(* CODESYS project beveling.project

Project tree, tasks and I/O mapping:
  Device : AM523-0808TN, Shenzhen Inovance Control Technology, version 3.5.11.50
      settings: PersistentStartAdddr = 0; PersistentStartEndAddr = 524287; Mode = 1
    application Application
      libraries: Standard, * (System); CmpEventMgr, 3.5.8.0 (System); Component Manager, 3.5.9.0 (System); CmpApp, 3.5.11.0 (System); CmpIecTask, 3.5.9.0 (System); CmpHCMotion, 1.1.8.0 (Inovance)
      task MainTask (cyclic, interval 4 ms, priority 1) calls nothing
      task ETHERCAT1 (cyclic, interval 2000 µs, priority 0) calls ETHERCAT1.EtherCAT_Task, PLC_PRG
      01_Data/
        global variables GVL_Parameters
        global variables GVL_IO_Physical
        global variables GVL_Modbus
        global variables GVL_RealDevice
        global variables GVL_DeviceIds
        global variables GVL_Simulation
        global variables GVL_Interface
        global variables GVL_IO
      06_Simulation/
        function block FB_SimDevice [ST]
        function block FB_SimPlant [ST]
      program PLC_PRG [ST]
      global variables GVL_Motion
      04_Machine/
        function block FB_IOMap [ST]
        function block FB_AlarmManager [ST]
        function block FB_PanelInput [ST]
        function block FB_AutoCycle [ST]
        function block FB_Interlocks [ST]
        function F_RecipeValid [ST]
        function block FB_ManualControl [ST]
        function block FB_Machine [ST]
        function block FB_Indicator [ST]
      00_Types/
        data type ST_RealDeviceSettings
        data type ST_MachineStatus
        data type E_MachineMode
        data type ST_Recipe
        data type ST_DeviceStatus
        data type E_DeviceAction
        data type E_MachineState
        data type ST_DeviceCommand
        data type ST_OperatorCommand
        data type ST_DeviceConfig
        data type ST_SimulationSettings
        data type E_DeviceKind
        data type ST_ManualCommand
        data type E_AutoStep
        data type ST_RemoteCommand
        data type ST_PanelInputs
      90_Legacy/
        program PRG_AxisDemo [ST]
      TaskEventPreStart
      05_Communication/
        function block FB_ModbusInterface [ST]
      03_Units/
        function block FB_ReturnKnife [ST]
        function block FB_PostCut [ST]
        function block FB_ResetLength [ST]
        function block FB_Initialize [ST]
        function block FB_Unload [ST]
        function block FB_ClearLength [ST]
        function block FB_ClearanceUnit [ST]
        function block FB_ClearTransfer [ST]
      DifferentialMonitor
      02_Devices/
        function block FB_RealAxis [ST]
        function block FB_RealCylinder [ST]
        function block FB_Motor [ST]
        function block FB_RealCylinderGroup [ST]
        function F_Done [ST]
        function block FB_Valve [ST]
        function F_At [ST]
        function block FB_Axis [ST]
        function F_SafetyBypassActive [ST]
        function block FB_RealSensor [ST]
        function block FB_Cylinder [ST]
        function F_Command [ST]
        function F_NextID [ST]
        function block FB_DeviceManager [ST]
    Device Diagnosis
    HardWare Configuration
    ConfigStorage
    Network Configuration
      LocalBus Config
      EtherCAT Config
    Resources List
    Serial : 串行接口, 汇川技术股份有限公司, version 00.00.00.10
      COM : Serial Port, Inovance, version 00.00.00.10
          settings: Device = AM523-0808TN; devGuid = 'e48f0cf2-85a4-455f-a8e7-135d3403221f'
    Local Bus
      GL20_0032ETN : GL20(GL20S) 32点DO模块, Inovance, version 00.00.00.10
          settings: ModuleBaseInfoStruct.BusType = 10; ModuleBaseInfoStruct.RackNumber = 1; ModuleBaseInfoStruct.SlotNumber = 2
          output Application.xDoG9Valve : BOOL  // QB(I).Q0
          output Application.xDoG1ValveL : BOOL  // QB(I).Q1
          output Application.xDoG1ValveR : BOOL  // QB(I).Q2
          output Application.xDoLampGreen : BOOL  // QB(II).Q0
          output Application.xDoLampRed : BOOL  // QB(II).Q1
          unmapped channels: QB(I), QB(II), QB(III), QB(IV)
      GL20_3200END : GL20(GL20S) 32通道DI模块, Inovance, version 00.00.00.10
          settings: ModuleBaseInfoStruct.BusType = 10; ModuleBaseInfoStruct.RackNumber = 1; ModuleBaseInfoStruct.SlotNumber = 1
          input  Application.xDiG1LRetract : BOOL  // IB(I).I0
          input  Application.xDiG1LExtend : BOOL  // IB(I).I1
          input  Application.xDiG1RRetract : BOOL  // IB(I).I2
          input  Application.xDiG1RExtend : BOOL  // IB(I).I3
          input  Application.xDiG9Retract : BOOL  // IB(I).I4
          input  Application.xDiG9Extend : BOOL  // IB(I).I5
          input  Application.xDiEStop : BOOL  // IB(II).I0
          input  Application.xDiPanelRunStop : BOOL  // IB(II).I1
          input  Application.xDiPanelStart : BOOL  // IB(II).I2
          input  Application.xDiPanelReset : BOOL  // IB(II).I3
          input  Application.xDiPanelInit : BOOL  // IB(II).I4
          input  Application.xDiPanelRunStart : BOOL  // IB(II).I5
          input  Application.xDiPanelAutoMode : BOOL  // IB(II).I6
          input  Application.xDiPanelSafetyPermit : BOOL  // IB(II).I7
          input  Application.xDiMaterialLength : BOOL  // IB(III).I0
          unmapped channels: IB(I), IB(II), IB(III), IB(IV)
    EXP_A : 扩展卡, 汇川技术股份有限公司, version 00.00.00.10
    ETHERCAT1 : EtherCAT Master SoftMotion, 3S - Smart Software Solutions GmbH, version 3.5.11.10
        settings:  = 0; MasterCycleTime = 2000; NetworkName = 'eth1'; SelectNetworkByName = TRUE; DisableTaskGeneration = True; SlaveArrayName = ADR(_EC1_Node)
      ASDA_B3_E_CoE_Drive_4 : Delta ASDA-B3-E EtherCAT(CoE) Drive, Delta Electronics, Inc., order no. ASDA-B3-E CoE Drive, version Revision=16#00030000
          settings: StationAlias = 0; Ring of slave = 0; Configuration address of the slave = 5; DC sync0 cycletime = 2000; DC sync1 cycletime = 2000; Interpolation time period.Value = 2
          unmapped channels: Control Word, Target Position, Target Velocity, Target Torque, Touch Probe Function, Status Word, Actual Position, Velocity actual value, Actual Torque, Touch Probe Status, Touch Probe Pos1 Pos Value, Digital inputs
        cetui : Axis, Inovance, order no. 0, version 4.0.0.0
            settings: wDriveID = 5; dwRatioTechUnitsDenom = 8388608; iRatioTechUnitsNum = 5; HomingMode = 2; ZeroSignal = 0; StartDirction = -1; EndDirection = -1; PosLimitMode = 1; NegLimitMode = 1; HomingVelocity = 30; HomingApproachVelocity = 10; HomingAcceleration = 100; HomingDeceleration = 100; HomingJerk = 0; HomeMaskDistance = 0; HomePositionOffset = 0; HomePushTime = 0; HomeCompensation = 0; HomeTimeout = 0; HomeCompensationVelocity = 1000; 4000 = 1; 4001 = 1; ScalingIncs = 16777216; ScalingGearOutput1 = 10; 6005 = 1; AdrOffset_8010 = 72; BitOffset_8010 = 0; BitLength_8010 = 16; Address_8010 = '%QW36'; Type_8010 = 'UINT'; AddressPointer_8010 = ADR(%QW36); AdrOffset_8020 = 76; BitOffset_8020 = 0; BitLength_8020 = 32; Address_8020 = '%QD19'; Type_8020 = 'DINT'; AddressPointer_8020 = ADR(%QD19); AdrOffset_8030 = 80; BitOffset_8030 = 0; BitLength_8030 = 32;
              Address_8030 = '%QD20'; Type_8030 = 'DINT'; AddressPointer_8030 = ADR(%QD20); AdrOffset_8040 = 84; BitOffset_8040 = 0; BitLength_8040 = 16; Address_8040 = '%QW42'; Type_8040 = 'INT'; AddressPointer_8040 = ADR(%QW42); AdrOffset_8050 = 4294967295; BitOffset_8050 = 0; BitLength_8050 = 0; Address_8050 = ''; Type_8050 = ''; AddressPointer_8050 = 0; AdrOffset_8060 = 86; BitOffset_8060 = 0; BitLength_8060 = 16; Address_8060 = '%QW43'; Type_8060 = 'UINT'; AddressPointer_8060 = ADR(%QW43); AdrOffset_8070 = 4294967295; BitOffset_8070 = 0; BitLength_8070 = 0; Address_8070 = ''; Type_8070 = ''; AddressPointer_8070 = 0; AdrOffset_8080 = 4294967295; BitOffset_8080 = 0; BitLength_8080 = 0; Address_8080 = ''; Type_8080 = ''; AddressPointer_8080 = 0; AdrOffset_8090 = 4294967295; BitOffset_8090 = 0; BitLength_8090 = 0; Address_8090 = ''; Type_8090 = ''; AddressPointer_8090 = 0; AdrOffset_8100 = 4294967295;
              BitOffset_8100 = 0; BitLength_8100 = 0; Address_8100 = ''; Type_8100 = ''; AddressPointer_8100 = 0; AdrOffset_8510 = 104; BitOffset_8510 = 0; BitLength_8510 = 16; Address_8510 = '%IW52'; Type_8510 = 'UINT'; AddressPointer_8510 = ADR(%IW52); AdrOffset_8520 = 108; BitOffset_8520 = 0; BitLength_8520 = 32; Address_8520 = '%ID27'; Type_8520 = 'DINT'; AddressPointer_8520 = ADR(%ID27); AdrOffset_8530 = 112; BitOffset_8530 = 0; BitLength_8530 = 32; Address_8530 = '%ID28'; Type_8530 = 'DINT'; AddressPointer_8530 = ADR(%ID28); AdrOffset_8540 = 116; BitOffset_8540 = 0; BitLength_8540 = 16; Address_8540 = '%IW58'; Type_8540 = 'INT'; AddressPointer_8540 = ADR(%IW58); AdrOffset_8550 = 4294967295; BitOffset_8550 = 0; BitLength_8550 = 0; Address_8550 = ''; Type_8550 = ''; AddressPointer_8550 = 0; AdrOffset_8560 = 124; BitOffset_8560 = 0; BitLength_8560 = 32; Address_8560 = '%ID31'; Type_8560 = 'UDINT';
              AddressPointer_8560 = ADR(%ID31); AdrOffset_8570 = 118; BitOffset_8570 = 0; BitLength_8570 = 16; Address_8570 = '%IW59'; Type_8570 = 'UINT'; AddressPointer_8570 = ADR(%IW59); AdrOffset_8580 = 120; BitOffset_8580 = 0; BitLength_8580 = 32; Address_8580 = '%ID30'; Type_8580 = 'DINT'; AddressPointer_8580 = ADR(%ID30); AdrOffset_8590 = 4294967295; BitOffset_8590 = 0; BitLength_8590 = 0; Address_8590 = ''; Type_8590 = ''; AddressPointer_8590 = 0; AdrOffset_8600 = 4294967295; BitOffset_8600 = 0; BitLength_8600 = 0; Address_8600 = ''; Type_8600 = ''; AddressPointer_8600 = 0; AdrOffset_8600 = 4294967295; BitOffset_8600 = 0; BitLength_8600 = 0; Address_8610 = ''; Type_8610 = ''; AddressPointer_8610 = 0; AdrOffset_8620 = 4294967295; BitOffset_8620 = 0; BitLength_8620 = 0; Address_8620 = ''; Type_8620 = ''; AddressPointer_8620 = 0; IsValid = True; AxisNumber = 5; IsHostHoming = True;
              PulseSelectIndex = 0
      DM3B_EC542 : DM3B-EC542(COE), Leadshine Technology Co.,Ltd., order no. DM3B-EC542, version Revision=16#00000001
          settings: StationAlias = 0; Ring of slave = 0; Configuration address of the slave = 8; DC sync0 cycletime = 2000; DC sync1 cycletime = 2000
          unmapped channels: Control Word, Profile Target Position, Touch Probe Function, Last Error Code, Status Word, Modes of Operation display, Position Actual Value, Touch Probe Status, Touch Probe 1 Positive Value, Digital Inputs
        dingchang_shangxia : Axis, Inovance, order no. 0, version 4.0.0.0
            settings: wDriveID = 8; dwRatioTechUnitsDenom = 10000; HomingMode = 7; ZeroSignal = 0; StartDirction = -1; EndDirection = 1; PosLimitMode = 0; NegLimitMode = 0; HomingVelocity = 5; HomingApproachVelocity = 2; HomingAcceleration = 100; HomingDeceleration = 100; HomingJerk = 0; HomeMaskDistance = 0; HomePositionOffset = 0; HomePushTime = 0; HomeCompensation = 0; HomeTimeout = 0; HomeCompensationVelocity = 1000; 4000 = 1; 4001 = 0; ScalingIncs = 10000; 6005 = 1; AdrOffset_8010 = 116; BitOffset_8010 = 0; BitLength_8010 = 16; Address_8010 = '%QW58'; Type_8010 = 'UINT'; AddressPointer_8010 = ADR(%QW58); AdrOffset_8020 = 120; BitOffset_8020 = 0; BitLength_8020 = 32; Address_8020 = '%QD30'; Type_8020 = 'DINT'; AddressPointer_8020 = ADR(%QD30); AdrOffset_8030 = 4294967295; BitOffset_8030 = 0; BitLength_8030 = 0; Address_8030 = ''; Type_8030 = '';
              AddressPointer_8030 = 0; AdrOffset_8040 = 4294967295; BitOffset_8040 = 0; BitLength_8040 = 0; Address_8040 = ''; Type_8040 = ''; AddressPointer_8040 = 0; AdrOffset_8050 = 4294967295; BitOffset_8050 = 0; BitLength_8050 = 0; Address_8050 = ''; Type_8050 = ''; AddressPointer_8050 = 0; AdrOffset_8060 = 124; BitOffset_8060 = 0; BitLength_8060 = 16; Address_8060 = '%QW62'; Type_8060 = 'UINT'; AddressPointer_8060 = ADR(%QW62); AdrOffset_8070 = 4294967295; BitOffset_8070 = 0; BitLength_8070 = 0; Address_8070 = ''; Type_8070 = ''; AddressPointer_8070 = 0; AdrOffset_8080 = 4294967295; BitOffset_8080 = 0; BitLength_8080 = 0; Address_8080 = ''; Type_8080 = ''; AddressPointer_8080 = 0; AdrOffset_8090 = 4294967295; BitOffset_8090 = 0; BitLength_8090 = 0; Address_8090 = ''; Type_8090 = ''; AddressPointer_8090 = 0; AdrOffset_8100 = 4294967295; BitOffset_8100 = 0; BitLength_8100 = 0;
              Address_8100 = ''; Type_8100 = ''; AddressPointer_8100 = 0; AdrOffset_8510 = 186; BitOffset_8510 = 0; BitLength_8510 = 16; Address_8510 = '%IW93'; Type_8510 = 'UINT'; AddressPointer_8510 = ADR(%IW93); AdrOffset_8520 = 192; BitOffset_8520 = 0; BitLength_8520 = 32; Address_8520 = '%ID48'; Type_8520 = 'DINT'; AddressPointer_8520 = ADR(%ID48); AdrOffset_8530 = 4294967295; BitOffset_8530 = 0; BitLength_8530 = 0; Address_8530 = ''; Type_8530 = ''; AddressPointer_8530 = 0; AdrOffset_8540 = 4294967295; BitOffset_8540 = 0; BitLength_8540 = 0; Address_8540 = ''; Type_8540 = ''; AddressPointer_8540 = 0; AdrOffset_8550 = 188; BitOffset_8550 = 0; BitLength_8550 = 8; Address_8550 = '%IB188'; Type_8550 = 'SINT'; AddressPointer_8550 = ADR(%IB188); AdrOffset_8560 = 204; BitOffset_8560 = 0; BitLength_8560 = 32; Address_8560 = '%ID51'; Type_8560 = 'UDINT'; AddressPointer_8560 = ADR(%ID51); AdrOffset_8570 = 196;
              BitOffset_8570 = 0; BitLength_8570 = 16; Address_8570 = '%IW98'; Type_8570 = 'UINT'; AddressPointer_8570 = ADR(%IW98); AdrOffset_8580 = 200; BitOffset_8580 = 0; BitLength_8580 = 32; Address_8580 = '%ID50'; Type_8580 = 'DINT'; AddressPointer_8580 = ADR(%ID50); AdrOffset_8590 = 4294967295; BitOffset_8590 = 0; BitLength_8590 = 0; Address_8590 = ''; Type_8590 = ''; AddressPointer_8590 = 0; AdrOffset_8600 = 4294967295; BitOffset_8600 = 0; BitLength_8600 = 0; Address_8600 = ''; Type_8600 = ''; AddressPointer_8600 = 0; AdrOffset_8600 = 4294967295; BitOffset_8600 = 0; BitLength_8600 = 0; Address_8610 = ''; Type_8610 = ''; AddressPointer_8610 = 0; AdrOffset_8620 = 184; BitOffset_8620 = 0; BitLength_8620 = 16; Address_8620 = '%IW92'; Type_8620 = 'UINT'; AddressPointer_8620 = ADR(%IW92); IsValid = True; AxisNumber = 8; IsHostHoming = True; PulseSelectIndex = 0
      ASDA_B3_E_CoE_Drive_1 : Delta ASDA-B3-E EtherCAT(CoE) Drive, Delta Electronics, Inc., order no. ASDA-B3-E CoE Drive, version Revision=16#00030000
          settings: StationAlias = 0; Ring of slave = 0; Configuration address of the slave = 1; DC sync0 cycletime = 2000; DC sync1 cycletime = 2000; Interpolation time period.Value = 2
          unmapped channels: Control Word, Target Position, Target Velocity, Target Torque, Touch Probe Function, Status Word, Actual Position, Velocity actual value, Actual Torque, Touch Probe Status, Touch Probe Pos1 Pos Value, Digital inputs
        qiege : Axis, Inovance, order no. 0, version 4.0.0.0
            settings: wDriveID = 2; dwRatioTechUnitsDenom = 4194304; iRatioTechUnitsNum = 5; HomingMode = 2; ZeroSignal = 0; StartDirction = -1; EndDirection = -1; PosLimitMode = 1; NegLimitMode = 1; HomingVelocity = 40; HomingApproachVelocity = 2; HomingAcceleration = 100; HomingDeceleration = 200; HomingJerk = 0; HomeMaskDistance = 0; HomePositionOffset = 0; HomePushTime = 0; HomeCompensation = 0; HomeTimeout = 0; HomeCompensationVelocity = 1000; 4000 = 1; 4001 = 1; ScalingIncs = 16777216; ScalingMotorTurns2 = 12; 6005 = 240; AdrOffset_8010 = 8; BitOffset_8010 = 0; BitLength_8010 = 16; Address_8010 = '%QW4'; Type_8010 = 'UINT'; AddressPointer_8010 = ADR(%QW4); AdrOffset_8020 = 12; BitOffset_8020 = 0; BitLength_8020 = 32; Address_8020 = '%QD3'; Type_8020 = 'DINT'; AddressPointer_8020 = ADR(%QD3); AdrOffset_8030 = 16; BitOffset_8030 = 0; BitLength_8030 = 32;
              Address_8030 = '%QD4'; Type_8030 = 'DINT'; AddressPointer_8030 = ADR(%QD4); AdrOffset_8040 = 20; BitOffset_8040 = 0; BitLength_8040 = 16; Address_8040 = '%QW10'; Type_8040 = 'INT'; AddressPointer_8040 = ADR(%QW10); AdrOffset_8050 = 4294967295; BitOffset_8050 = 0; BitLength_8050 = 0; Address_8050 = ''; Type_8050 = ''; AddressPointer_8050 = 0; AdrOffset_8060 = 22; BitOffset_8060 = 0; BitLength_8060 = 16; Address_8060 = '%QW11'; Type_8060 = 'UINT'; AddressPointer_8060 = ADR(%QW11); AdrOffset_8070 = 4294967295; BitOffset_8070 = 0; BitLength_8070 = 0; Address_8070 = ''; Type_8070 = ''; AddressPointer_8070 = 0; AdrOffset_8080 = 4294967295; BitOffset_8080 = 0; BitLength_8080 = 0; Address_8080 = ''; Type_8080 = ''; AddressPointer_8080 = 0; AdrOffset_8090 = 4294967295; BitOffset_8090 = 0; BitLength_8090 = 0; Address_8090 = ''; Type_8090 = ''; AddressPointer_8090 = 0; AdrOffset_8100 = 4294967295;
              BitOffset_8100 = 0; BitLength_8100 = 0; Address_8100 = ''; Type_8100 = ''; AddressPointer_8100 = 0; AdrOffset_8510 = 8; BitOffset_8510 = 0; BitLength_8510 = 16; Address_8510 = '%IW4'; Type_8510 = 'UINT'; AddressPointer_8510 = ADR(%IW4); AdrOffset_8520 = 12; BitOffset_8520 = 0; BitLength_8520 = 32; Address_8520 = '%ID3'; Type_8520 = 'DINT'; AddressPointer_8520 = ADR(%ID3); AdrOffset_8530 = 16; BitOffset_8530 = 0; BitLength_8530 = 32; Address_8530 = '%ID4'; Type_8530 = 'DINT'; AddressPointer_8530 = ADR(%ID4); AdrOffset_8540 = 20; BitOffset_8540 = 0; BitLength_8540 = 16; Address_8540 = '%IW10'; Type_8540 = 'INT'; AddressPointer_8540 = ADR(%IW10); AdrOffset_8550 = 4294967295; BitOffset_8550 = 0; BitLength_8550 = 0; Address_8550 = ''; Type_8550 = ''; AddressPointer_8550 = 0; AdrOffset_8560 = 28; BitOffset_8560 = 0; BitLength_8560 = 32; Address_8560 = '%ID7'; Type_8560 = 'UDINT';
              AddressPointer_8560 = ADR(%ID7); AdrOffset_8570 = 22; BitOffset_8570 = 0; BitLength_8570 = 16; Address_8570 = '%IW11'; Type_8570 = 'UINT'; AddressPointer_8570 = ADR(%IW11); AdrOffset_8580 = 24; BitOffset_8580 = 0; BitLength_8580 = 32; Address_8580 = '%ID6'; Type_8580 = 'DINT'; AddressPointer_8580 = ADR(%ID6); AdrOffset_8590 = 4294967295; BitOffset_8590 = 0; BitLength_8590 = 0; Address_8590 = ''; Type_8590 = ''; AddressPointer_8590 = 0; AdrOffset_8600 = 4294967295; BitOffset_8600 = 0; BitLength_8600 = 0; Address_8600 = ''; Type_8600 = ''; AddressPointer_8600 = 0; AdrOffset_8600 = 4294967295; BitOffset_8600 = 0; BitLength_8600 = 0; Address_8610 = ''; Type_8610 = ''; AddressPointer_8610 = 0; AdrOffset_8620 = 4294967295; BitOffset_8620 = 0; BitLength_8620 = 0; Address_8620 = ''; Type_8620 = ''; AddressPointer_8620 = 0; IsValid = True; AxisNumber = 1; IsHostHoming = True;
              PulseSelectIndex = 0
      ASDA_B3_E_CoE_Drive_5 : Delta ASDA-B3-E EtherCAT(CoE) Drive, Delta Electronics, Inc., order no. ASDA-B3-E CoE Drive, version Revision=16#00030000
          settings: StationAlias = 0; Ring of slave = 0; Configuration address of the slave = 7; DC sync0 cycletime = 2000; DC sync1 cycletime = 2000; Interpolation time period.Value = 2
          unmapped channels: Control Word, Target Position, Target Velocity, Target Torque, Touch Probe Function, Status Word, Actual Position, Velocity actual value, Actual Torque, Touch Probe Status, Touch Probe Pos1 Pos Value, Digital inputs
        jixieshou : Axis, Inovance, order no. 0, version 4.0.0.0
            settings: wDriveID = 7; dwRatioTechUnitsDenom = 10485760; HomingMode = 10; ZeroSignal = 0; StartDirction = 1; EndDirection = 1; PosLimitMode = 0; NegLimitMode = 0; HomingVelocity = 10; HomingApproachVelocity = 2; HomingAcceleration = 100; HomingDeceleration = 100; HomingJerk = 0; HomeMaskDistance = 0; HomePositionOffset = 0; HomePushTime = 0; HomeCompensation = 0; HomeTimeout = 0; HomeCompensationVelocity = 1000; 4000 = 1; 4001 = 1; ScalingIncs = 16777216; ScalingMotorTurns2 = 10; ScalingGearOutput1 = 16; 6005 = 1; AdrOffset_8010 = 100; BitOffset_8010 = 0; BitLength_8010 = 16; Address_8010 = '%QW50'; Type_8010 = 'UINT'; AddressPointer_8010 = ADR(%QW50); AdrOffset_8020 = 104; BitOffset_8020 = 0; BitLength_8020 = 32; Address_8020 = '%QD26'; Type_8020 = 'DINT'; AddressPointer_8020 = ADR(%QD26); AdrOffset_8030 = 108; BitOffset_8030 = 0; BitLength_8030 = 32;
              Address_8030 = '%QD27'; Type_8030 = 'DINT'; AddressPointer_8030 = ADR(%QD27); AdrOffset_8040 = 112; BitOffset_8040 = 0; BitLength_8040 = 16; Address_8040 = '%QW56'; Type_8040 = 'INT'; AddressPointer_8040 = ADR(%QW56); AdrOffset_8050 = 4294967295; BitOffset_8050 = 0; BitLength_8050 = 0; Address_8050 = ''; Type_8050 = ''; AddressPointer_8050 = 0; AdrOffset_8060 = 114; BitOffset_8060 = 0; BitLength_8060 = 16; Address_8060 = '%QW57'; Type_8060 = 'UINT'; AddressPointer_8060 = ADR(%QW57); AdrOffset_8070 = 4294967295; BitOffset_8070 = 0; BitLength_8070 = 0; Address_8070 = ''; Type_8070 = ''; AddressPointer_8070 = 0; AdrOffset_8080 = 4294967295; BitOffset_8080 = 0; BitLength_8080 = 0; Address_8080 = ''; Type_8080 = ''; AddressPointer_8080 = 0; AdrOffset_8090 = 4294967295; BitOffset_8090 = 0; BitLength_8090 = 0; Address_8090 = ''; Type_8090 = ''; AddressPointer_8090 = 0; AdrOffset_8100 = 4294967295;
              BitOffset_8100 = 0; BitLength_8100 = 0; Address_8100 = ''; Type_8100 = ''; AddressPointer_8100 = 0; AdrOffset_8510 = 160; BitOffset_8510 = 0; BitLength_8510 = 16; Address_8510 = '%IW80'; Type_8510 = 'UINT'; AddressPointer_8510 = ADR(%IW80); AdrOffset_8520 = 164; BitOffset_8520 = 0; BitLength_8520 = 32; Address_8520 = '%ID41'; Type_8520 = 'DINT'; AddressPointer_8520 = ADR(%ID41); AdrOffset_8530 = 168; BitOffset_8530 = 0; BitLength_8530 = 32; Address_8530 = '%ID42'; Type_8530 = 'DINT'; AddressPointer_8530 = ADR(%ID42); AdrOffset_8540 = 172; BitOffset_8540 = 0; BitLength_8540 = 16; Address_8540 = '%IW86'; Type_8540 = 'INT'; AddressPointer_8540 = ADR(%IW86); AdrOffset_8550 = 4294967295; BitOffset_8550 = 0; BitLength_8550 = 0; Address_8550 = ''; Type_8550 = ''; AddressPointer_8550 = 0; AdrOffset_8560 = 180; BitOffset_8560 = 0; BitLength_8560 = 32; Address_8560 = '%ID45'; Type_8560 = 'UDINT';
              AddressPointer_8560 = ADR(%ID45); AdrOffset_8570 = 174; BitOffset_8570 = 0; BitLength_8570 = 16; Address_8570 = '%IW87'; Type_8570 = 'UINT'; AddressPointer_8570 = ADR(%IW87); AdrOffset_8580 = 176; BitOffset_8580 = 0; BitLength_8580 = 32; Address_8580 = '%ID44'; Type_8580 = 'DINT'; AddressPointer_8580 = ADR(%ID44); AdrOffset_8590 = 4294967295; BitOffset_8590 = 0; BitLength_8590 = 0; Address_8590 = ''; Type_8590 = ''; AddressPointer_8590 = 0; AdrOffset_8600 = 4294967295; BitOffset_8600 = 0; BitLength_8600 = 0; Address_8600 = ''; Type_8600 = ''; AddressPointer_8600 = 0; AdrOffset_8600 = 4294967295; BitOffset_8600 = 0; BitLength_8600 = 0; Address_8610 = ''; Type_8610 = ''; AddressPointer_8610 = 0; AdrOffset_8620 = 4294967295; BitOffset_8620 = 0; BitLength_8620 = 0; Address_8620 = ''; Type_8620 = ''; AddressPointer_8620 = 0; IsValid = True; AxisNumber = 7; IsHostHoming = True;
              PulseSelectIndex = 0
      ASDA_B3_E_CoE_Drive : Delta ASDA-B3-E EtherCAT(CoE) Drive, Delta Electronics, Inc., order no. ASDA-B3-E CoE Drive, version Revision=16#00030000
          settings: StationAlias = 0; Ring of slave = 0; Configuration address of the slave = 2; AutoUpdate = False; DC sync0 cycletime = 2000; DC sync0 cycletime = 2000000; DC sync1 cycletime = 2000; DC sync1 cycletime = 2000000; DC sync1 factor = 'x 1'; Interpolation time period.Value = 2
          unmapped channels: Control Word, Target Position, Target Velocity, Target Torque, Touch Probe Function, Status Word, Actual Position, Velocity actual value, Actual Torque, Touch Probe Status, Touch Probe Pos1 Pos Value, Digital inputs
        xuanzhuan : Axis, Inovance, order no. 0, version 4.0.0.0
            settings: dwRatioTechUnitsDenom = 45088768; iRatioTechUnitsNum = 9; iMovementType = 0; fSWMaxVelocity = 10; fSWMaxAcceleration = 100; fSWMaxDeceleration = 100; HomingMode = 2; ZeroSignal = 0; StartDirction = -1; EndDirection = -1; PosLimitMode = 1; NegLimitMode = 1; HomingVelocity = 3; HomingApproachVelocity = 1; HomingAcceleration = 100; HomingDeceleration = 100; HomingJerk = 0; HomeMaskDistance = 0; HomePositionOffset = 0; HomePushTime = 0; HomeCompensation = 0; HomeTimeout = 0; HomeCompensationVelocity = 1000; 4000 = 4; 4001 = 1; ScalingIncs = 16777216; ScalingMotorTurns2 = 215; ScalingGearOutput1 = 2; 6005 = 360; AdrOffset_8010 = 24; BitOffset_8010 = 0; BitLength_8010 = 16; Address_8010 = '%QW12'; Type_8010 = 'UINT'; AddressPointer_8010 = ADR(%QW12); AdrOffset_8020 = 28; BitOffset_8020 = 0; BitLength_8020 = 32; Address_8020 = '%QD7'; Type_8020 = 'DINT';
              AddressPointer_8020 = ADR(%QD7); AdrOffset_8030 = 32; BitOffset_8030 = 0; BitLength_8030 = 32; Address_8030 = '%QD8'; Type_8030 = 'DINT'; AddressPointer_8030 = ADR(%QD8); AdrOffset_8040 = 36; BitOffset_8040 = 0; BitLength_8040 = 16; Address_8040 = '%QW18'; Type_8040 = 'INT'; AddressPointer_8040 = ADR(%QW18); AdrOffset_8050 = 4294967295; BitOffset_8050 = 0; BitLength_8050 = 0; Address_8050 = ''; Type_8050 = ''; AddressPointer_8050 = 0; AdrOffset_8060 = 38; BitOffset_8060 = 0; BitLength_8060 = 16; Address_8060 = '%QW19'; Type_8060 = 'UINT'; AddressPointer_8060 = ADR(%QW19); AdrOffset_8070 = 4294967295; BitOffset_8070 = 0; BitLength_8070 = 0; Address_8070 = ''; Type_8070 = ''; AddressPointer_8070 = 0; AdrOffset_8080 = 4294967295; BitOffset_8080 = 0; BitLength_8080 = 0; Address_8080 = ''; Type_8080 = ''; AddressPointer_8080 = 0; AdrOffset_8090 = 4294967295; BitOffset_8090 = 0; BitLength_8090 = 0;
              Address_8090 = ''; Type_8090 = ''; AddressPointer_8090 = 0; AdrOffset_8100 = 4294967295; BitOffset_8100 = 0; BitLength_8100 = 0; Address_8100 = ''; Type_8100 = ''; AddressPointer_8100 = 0; AdrOffset_8510 = 32; BitOffset_8510 = 0; BitLength_8510 = 16; Address_8510 = '%IW16'; Type_8510 = 'UINT'; AddressPointer_8510 = ADR(%IW16); AdrOffset_8520 = 36; BitOffset_8520 = 0; BitLength_8520 = 32; Address_8520 = '%ID9'; Type_8520 = 'DINT'; AddressPointer_8520 = ADR(%ID9); AdrOffset_8530 = 40; BitOffset_8530 = 0; BitLength_8530 = 32; Address_8530 = '%ID10'; Type_8530 = 'DINT'; AddressPointer_8530 = ADR(%ID10); AdrOffset_8540 = 44; BitOffset_8540 = 0; BitLength_8540 = 16; Address_8540 = '%IW22'; Type_8540 = 'INT'; AddressPointer_8540 = ADR(%IW22); AdrOffset_8550 = 4294967295; BitOffset_8550 = 0; BitLength_8550 = 0; Address_8550 = ''; Type_8550 = ''; AddressPointer_8550 = 0; AdrOffset_8560 = 52;
              BitOffset_8560 = 0; BitLength_8560 = 32; Address_8560 = '%ID13'; Type_8560 = 'UDINT'; AddressPointer_8560 = ADR(%ID13); AdrOffset_8570 = 46; BitOffset_8570 = 0; BitLength_8570 = 16; Address_8570 = '%IW23'; Type_8570 = 'UINT'; AddressPointer_8570 = ADR(%IW23); AdrOffset_8580 = 48; BitOffset_8580 = 0; BitLength_8580 = 32; Address_8580 = '%ID12'; Type_8580 = 'DINT'; AddressPointer_8580 = ADR(%ID12); AdrOffset_8590 = 4294967295; BitOffset_8590 = 0; BitLength_8590 = 0; Address_8590 = ''; Type_8590 = ''; AddressPointer_8590 = 0; AdrOffset_8600 = 4294967295; BitOffset_8600 = 0; BitLength_8600 = 0; Address_8600 = ''; Type_8600 = ''; AddressPointer_8600 = 0; AdrOffset_8600 = 4294967295; BitOffset_8600 = 0; BitLength_8600 = 0; Address_8610 = ''; Type_8610 = ''; AddressPointer_8610 = 0; AdrOffset_8620 = 4294967295; BitOffset_8620 = 0; BitLength_8620 = 0; Address_8620 = ''; Type_8620 = '';
              AddressPointer_8620 = 0; IsValid = True; AxisNumber = 2; IsHostHoming = True; PulseSelectIndex = 0
      HD3_EL : HD3_EL_V1.0, HUACHUANG, order no. HD3_EL, version Revision=16#00010001
          settings: StationAlias = 0; Ring of slave = 0; Configuration address of the slave = 6; AutoUpdate = False; DC sync0 cycletime = 2000; DC sync1 cycletime = 2000
          unmapped channels: Controlword, Target position, Touch probe function, Statusword, Position actual value, Touch probe status, Touch probe pos1 pos value, Touch probe pos2 pos value, Error code, Digital inputs, Modes of operation display
        dingchang_zuoyou : Axis, Inovance, order no. 0, version 4.0.0.0
            settings: wDriveID = 6; dwRatioTechUnitsDenom = 1000; HomingMode = 2; ZeroSignal = 0; StartDirction = -1; EndDirection = -1; PosLimitMode = 1; NegLimitMode = 1; HomingVelocity = 30; HomingApproachVelocity = 10; HomingAcceleration = 100; HomingDeceleration = 100; HomingJerk = 0; HomeMaskDistance = 0; HomePositionOffset = 0; HomePushTime = 0; HomeCompensation = 0; HomeTimeout = 0; HomeCompensationVelocity = 1000; 4000 = 1; 4001 = 0; ScalingIncs = 1000; 6005 = 1; AdrOffset_8010 = 88; BitOffset_8010 = 0; BitLength_8010 = 16; Address_8010 = '%QW44'; Type_8010 = 'UINT'; AddressPointer_8010 = ADR(%QW44); AdrOffset_8020 = 92; BitOffset_8020 = 0; BitLength_8020 = 32; Address_8020 = '%QD23'; Type_8020 = 'DINT'; AddressPointer_8020 = ADR(%QD23); AdrOffset_8030 = 4294967295; BitOffset_8030 = 0; BitLength_8030 = 0; Address_8030 = ''; Type_8030 = '';
              AddressPointer_8030 = 0; AdrOffset_8040 = 4294967295; BitOffset_8040 = 0; BitLength_8040 = 0; Address_8040 = ''; Type_8040 = ''; AddressPointer_8040 = 0; AdrOffset_8050 = 4294967295; BitOffset_8050 = 0; BitLength_8050 = 0; Address_8050 = ''; Type_8050 = ''; AddressPointer_8050 = 0; AdrOffset_8060 = 96; BitOffset_8060 = 0; BitLength_8060 = 16; Address_8060 = '%QW48'; Type_8060 = 'UINT'; AddressPointer_8060 = ADR(%QW48); AdrOffset_8070 = 4294967295; BitOffset_8070 = 0; BitLength_8070 = 0; Address_8070 = ''; Type_8070 = ''; AddressPointer_8070 = 0; AdrOffset_8080 = 4294967295; BitOffset_8080 = 0; BitLength_8080 = 0; Address_8080 = ''; Type_8080 = ''; AddressPointer_8080 = 0; AdrOffset_8090 = 4294967295; BitOffset_8090 = 0; BitLength_8090 = 0; Address_8090 = ''; Type_8090 = ''; AddressPointer_8090 = 0; AdrOffset_8100 = 4294967295; BitOffset_8100 = 0; BitLength_8100 = 0;
              Address_8100 = ''; Type_8100 = ''; AddressPointer_8100 = 0; AdrOffset_8510 = 128; BitOffset_8510 = 0; BitLength_8510 = 16; Address_8510 = '%IW64'; Type_8510 = 'UINT'; AddressPointer_8510 = ADR(%IW64); AdrOffset_8520 = 132; BitOffset_8520 = 0; BitLength_8520 = 32; Address_8520 = '%ID33'; Type_8520 = 'DINT'; AddressPointer_8520 = ADR(%ID33); AdrOffset_8530 = 4294967295; BitOffset_8530 = 0; BitLength_8530 = 0; Address_8530 = ''; Type_8530 = ''; AddressPointer_8530 = 0; AdrOffset_8540 = 4294967295; BitOffset_8540 = 0; BitLength_8540 = 0; Address_8540 = ''; Type_8540 = ''; AddressPointer_8540 = 0; AdrOffset_8550 = 156; BitOffset_8550 = 0; BitLength_8550 = 8; Address_8550 = '%IB156'; Type_8550 = 'SINT'; AddressPointer_8550 = ADR(%IB156); AdrOffset_8560 = 152; BitOffset_8560 = 0; BitLength_8560 = 32; Address_8560 = '%ID38'; Type_8560 = 'UDINT'; AddressPointer_8560 = ADR(%ID38); AdrOffset_8570 = 136;
              BitOffset_8570 = 0; BitLength_8570 = 16; Address_8570 = '%IW68'; Type_8570 = 'UINT'; AddressPointer_8570 = ADR(%IW68); AdrOffset_8580 = 140; BitOffset_8580 = 0; BitLength_8580 = 32; Address_8580 = '%ID35'; Type_8580 = 'DINT'; AddressPointer_8580 = ADR(%ID35); AdrOffset_8590 = 4294967295; BitOffset_8590 = 0; BitLength_8590 = 0; Address_8590 = ''; Type_8590 = ''; AddressPointer_8590 = 0; AdrOffset_8600 = 144; BitOffset_8600 = 0; BitLength_8600 = 32; Address_8600 = '%ID36'; Type_8600 = 'DINT'; AddressPointer_8600 = ADR(%ID36); AdrOffset_8600 = 4294967295; BitOffset_8600 = 0; BitLength_8600 = 0; Address_8610 = ''; Type_8610 = ''; AddressPointer_8610 = 0; AdrOffset_8620 = 148; BitOffset_8620 = 0; BitLength_8620 = 16; Address_8620 = '%IW74'; Type_8620 = 'UINT'; AddressPointer_8620 = ADR(%IW74); IsValid = True; AxisNumber = 6; IsHostHoming = True; PulseSelectIndex = 0
      ASDA_B3_E_CoE_Drive_2 : Delta ASDA-B3-E EtherCAT(CoE) Drive, Delta Electronics, Inc., order no. ASDA-B3-E CoE Drive, version Revision=16#00030000
          settings: StationAlias = 0; Ring of slave = 0; Configuration address of the slave = 3; DC sync0 cycletime = 2000; DC sync1 cycletime = 2000; Interpolation time period.Value = 2
          unmapped channels: Control Word, Target Position, Target Velocity, Target Torque, Touch Probe Function, Status Word, Actual Position, Velocity actual value, Actual Torque, Touch Probe Status, Touch Probe Pos1 Pos Value, Digital inputs
        pandao : Axis, Inovance, order no. 0, version 4.0.0.0
            settings: wDriveID = 3; dwRatioTechUnitsDenom = 16777216; HomingMode = 10; ZeroSignal = 0; StartDirction = 1; EndDirection = 1; PosLimitMode = 0; NegLimitMode = 0; HomingVelocity = 10; HomingApproachVelocity = 2; HomingAcceleration = 100; HomingDeceleration = 100; HomingJerk = 0; HomeMaskDistance = 0; HomePositionOffset = 0; HomePushTime = 0; HomeCompensation = 0; HomeTimeout = 0; HomeCompensationVelocity = 1000; 4000 = 0; 4001 = 0; ScalingIncs = 16777216; 6005 = 1; AdrOffset_8010 = 40; BitOffset_8010 = 0; BitLength_8010 = 16; Address_8010 = '%QW20'; Type_8010 = 'UINT'; AddressPointer_8010 = ADR(%QW20); AdrOffset_8020 = 44; BitOffset_8020 = 0; BitLength_8020 = 32; Address_8020 = '%QD11'; Type_8020 = 'DINT'; AddressPointer_8020 = ADR(%QD11); AdrOffset_8030 = 48; BitOffset_8030 = 0; BitLength_8030 = 32; Address_8030 = '%QD12'; Type_8030 = 'DINT';
              AddressPointer_8030 = ADR(%QD12); AdrOffset_8040 = 52; BitOffset_8040 = 0; BitLength_8040 = 16; Address_8040 = '%QW26'; Type_8040 = 'INT'; AddressPointer_8040 = ADR(%QW26); AdrOffset_8050 = 4294967295; BitOffset_8050 = 0; BitLength_8050 = 0; Address_8050 = ''; Type_8050 = ''; AddressPointer_8050 = 0; AdrOffset_8060 = 54; BitOffset_8060 = 0; BitLength_8060 = 16; Address_8060 = '%QW27'; Type_8060 = 'UINT'; AddressPointer_8060 = ADR(%QW27); AdrOffset_8070 = 4294967295; BitOffset_8070 = 0; BitLength_8070 = 0; Address_8070 = ''; Type_8070 = ''; AddressPointer_8070 = 0; AdrOffset_8080 = 4294967295; BitOffset_8080 = 0; BitLength_8080 = 0; Address_8080 = ''; Type_8080 = ''; AddressPointer_8080 = 0; AdrOffset_8090 = 4294967295; BitOffset_8090 = 0; BitLength_8090 = 0; Address_8090 = ''; Type_8090 = ''; AddressPointer_8090 = 0; AdrOffset_8100 = 4294967295; BitOffset_8100 = 0; BitLength_8100 = 0;
              Address_8100 = ''; Type_8100 = ''; AddressPointer_8100 = 0; AdrOffset_8510 = 56; BitOffset_8510 = 0; BitLength_8510 = 16; Address_8510 = '%IW28'; Type_8510 = 'UINT'; AddressPointer_8510 = ADR(%IW28); AdrOffset_8520 = 60; BitOffset_8520 = 0; BitLength_8520 = 32; Address_8520 = '%ID15'; Type_8520 = 'DINT'; AddressPointer_8520 = ADR(%ID15); AdrOffset_8530 = 64; BitOffset_8530 = 0; BitLength_8530 = 32; Address_8530 = '%ID16'; Type_8530 = 'DINT'; AddressPointer_8530 = ADR(%ID16); AdrOffset_8540 = 68; BitOffset_8540 = 0; BitLength_8540 = 16; Address_8540 = '%IW34'; Type_8540 = 'INT'; AddressPointer_8540 = ADR(%IW34); AdrOffset_8550 = 4294967295; BitOffset_8550 = 0; BitLength_8550 = 0; Address_8550 = ''; Type_8550 = ''; AddressPointer_8550 = 0; AdrOffset_8560 = 76; BitOffset_8560 = 0; BitLength_8560 = 32; Address_8560 = '%ID19'; Type_8560 = 'UDINT'; AddressPointer_8560 = ADR(%ID19); AdrOffset_8570 = 70;
              BitOffset_8570 = 0; BitLength_8570 = 16; Address_8570 = '%IW35'; Type_8570 = 'UINT'; AddressPointer_8570 = ADR(%IW35); AdrOffset_8580 = 72; BitOffset_8580 = 0; BitLength_8580 = 32; Address_8580 = '%ID18'; Type_8580 = 'DINT'; AddressPointer_8580 = ADR(%ID18); AdrOffset_8590 = 4294967295; BitOffset_8590 = 0; BitLength_8590 = 0; Address_8590 = ''; Type_8590 = ''; AddressPointer_8590 = 0; AdrOffset_8600 = 4294967295; BitOffset_8600 = 0; BitLength_8600 = 0; Address_8600 = ''; Type_8600 = ''; AddressPointer_8600 = 0; AdrOffset_8600 = 4294967295; BitOffset_8600 = 0; BitLength_8600 = 0; Address_8610 = ''; Type_8610 = ''; AddressPointer_8610 = 0; AdrOffset_8620 = 4294967295; BitOffset_8620 = 0; BitLength_8620 = 0; Address_8620 = ''; Type_8620 = ''; AddressPointer_8620 = 0; IsValid = True; AxisNumber = 3; IsHostHoming = True; PulseSelectIndex = 0
      ASDA_B3_E_CoE_Drive_3 : Delta ASDA-B3-E EtherCAT(CoE) Drive, Delta Electronics, Inc., order no. ASDA-B3-E CoE Drive, version Revision=16#00030000
          settings: StationAlias = 0; Ring of slave = 0; Configuration address of the slave = 4; DC sync0 cycletime = 2000; DC sync1 cycletime = 2000; Interpolation time period.Value = 2
          unmapped channels: Control Word, Target Position, Target Velocity, Target Torque, Touch Probe Function, Status Word, Actual Position, Velocity actual value, Actual Torque, Touch Probe Status, Touch Probe Pos1 Pos Value, Digital inputs
        songliao : Axis, Inovance, order no. 0, version 4.0.0.0
            settings: wDriveID = 4; dwRatioTechUnitsDenom = 3355443200; iRatioTechUnitsNum = 8231; fSWMaxVelocity = 50; fSWMaxAcceleration = 100; fSWMaxDeceleration = 100; fSWMaxJerk = 1000; HomingMode = 10; ZeroSignal = 0; StartDirction = 1; EndDirection = 1; PosLimitMode = 0; NegLimitMode = 0; HomingVelocity = 10; HomingApproachVelocity = 2; HomingAcceleration = 100; HomingDeceleration = 100; HomingJerk = 0; HomeMaskDistance = 0; HomePositionOffset = 0; HomePushTime = 0; HomeCompensation = 0; HomeTimeout = 0; HomeCompensationVelocity = 1000; 4000 = 1; 4001 = 1; ScalingIncs = 16777216; ScalingMotorTurns2 = 10; 6005 = 411.55; AdrOffset_8010 = 56; BitOffset_8010 = 0; BitLength_8010 = 16; Address_8010 = '%QW28'; Type_8010 = 'UINT'; AddressPointer_8010 = ADR(%QW28); AdrOffset_8020 = 60; BitOffset_8020 = 0; BitLength_8020 = 32; Address_8020 = '%QD15'; Type_8020 = 'DINT';
              AddressPointer_8020 = ADR(%QD15); AdrOffset_8030 = 64; BitOffset_8030 = 0; BitLength_8030 = 32; Address_8030 = '%QD16'; Type_8030 = 'DINT'; AddressPointer_8030 = ADR(%QD16); AdrOffset_8040 = 68; BitOffset_8040 = 0; BitLength_8040 = 16; Address_8040 = '%QW34'; Type_8040 = 'INT'; AddressPointer_8040 = ADR(%QW34); AdrOffset_8050 = 4294967295; BitOffset_8050 = 0; BitLength_8050 = 0; Address_8050 = ''; Type_8050 = ''; AddressPointer_8050 = 0; AdrOffset_8060 = 70; BitOffset_8060 = 0; BitLength_8060 = 16; Address_8060 = '%QW35'; Type_8060 = 'UINT'; AddressPointer_8060 = ADR(%QW35); AdrOffset_8070 = 4294967295; BitOffset_8070 = 0; BitLength_8070 = 0; Address_8070 = ''; Type_8070 = ''; AddressPointer_8070 = 0; AdrOffset_8080 = 4294967295; BitOffset_8080 = 0; BitLength_8080 = 0; Address_8080 = ''; Type_8080 = ''; AddressPointer_8080 = 0; AdrOffset_8090 = 4294967295; BitOffset_8090 = 0; BitLength_8090 = 0;
              Address_8090 = ''; Type_8090 = ''; AddressPointer_8090 = 0; AdrOffset_8100 = 4294967295; BitOffset_8100 = 0; BitLength_8100 = 0; Address_8100 = ''; Type_8100 = ''; AddressPointer_8100 = 0; AdrOffset_8510 = 80; BitOffset_8510 = 0; BitLength_8510 = 16; Address_8510 = '%IW40'; Type_8510 = 'UINT'; AddressPointer_8510 = ADR(%IW40); AdrOffset_8520 = 84; BitOffset_8520 = 0; BitLength_8520 = 32; Address_8520 = '%ID21'; Type_8520 = 'DINT'; AddressPointer_8520 = ADR(%ID21); AdrOffset_8530 = 88; BitOffset_8530 = 0; BitLength_8530 = 32; Address_8530 = '%ID22'; Type_8530 = 'DINT'; AddressPointer_8530 = ADR(%ID22); AdrOffset_8540 = 92; BitOffset_8540 = 0; BitLength_8540 = 16; Address_8540 = '%IW46'; Type_8540 = 'INT'; AddressPointer_8540 = ADR(%IW46); AdrOffset_8550 = 4294967295; BitOffset_8550 = 0; BitLength_8550 = 0; Address_8550 = ''; Type_8550 = ''; AddressPointer_8550 = 0; AdrOffset_8560 = 100;
              BitOffset_8560 = 0; BitLength_8560 = 32; Address_8560 = '%ID25'; Type_8560 = 'UDINT'; AddressPointer_8560 = ADR(%ID25); AdrOffset_8570 = 94; BitOffset_8570 = 0; BitLength_8570 = 16; Address_8570 = '%IW47'; Type_8570 = 'UINT'; AddressPointer_8570 = ADR(%IW47); AdrOffset_8580 = 96; BitOffset_8580 = 0; BitLength_8580 = 32; Address_8580 = '%ID24'; Type_8580 = 'DINT'; AddressPointer_8580 = ADR(%ID24); AdrOffset_8590 = 4294967295; BitOffset_8590 = 0; BitLength_8590 = 0; Address_8590 = ''; Type_8590 = ''; AddressPointer_8590 = 0; AdrOffset_8600 = 4294967295; BitOffset_8600 = 0; BitLength_8600 = 0; Address_8600 = ''; Type_8600 = ''; AddressPointer_8600 = 0; AdrOffset_8600 = 4294967295; BitOffset_8600 = 0; BitLength_8600 = 0; Address_8610 = ''; Type_8610 = ''; AddressPointer_8610 = 0; AdrOffset_8620 = 4294967295; BitOffset_8620 = 0; BitLength_8620 = 0; Address_8620 = ''; Type_8620 = '';
              AddressPointer_8620 = 0; IsValid = True; AxisNumber = 4; IsHostHoming = True; PulseSelectIndex = 0
    SoftMotion General Axis Pool
    EXP_B : 扩展卡, 汇川技术股份有限公司, version 00.00.00.10
    CAN : CAN总线, INOVANCE, version 00.00.00.10
    LocalHSIO : 本地高速IO, 汇川技术股份有限公司, version 2.0.0.0
        unmapped channels: %IB0 DigitalInput, %QB0 DigitalOutput
    HwConfiguratioinDevice : SystemConfig, Inovance, version 00.00.00.10
        settings: NetworkConfigArray.NetworkConfigArray.BusType = 10; NetworkConfigArray.NetworkConfigArray.RackSum = 1; NetworkConfigArray.NetworkConfigArray.HardwareConfigArray.HardwareConfigArray.RackNo = 1; NetworkConfigArray.NetworkConfigArray.HardwareConfigArray.HardwareConfigArray.ModuleNum = 2; EnableFun = 1
*)

// Device/Application/00_Types/ST_RealDeviceSettings
(* 模块说明：真实设备接管与调试旁路设置。默认接管 1、2、3、8、9、10、17 七台（现场已接线的轴与气缸），其余仍走仿真。 *)
TYPE ST_RealDeviceSettings :
STRUCT
axRealDevice : ARRAY[1..17] OF BOOL :=
    [TRUE, TRUE, TRUE, FALSE, FALSE, TRUE, FALSE, TRUE, TRUE, TRUE, FALSE, FALSE, FALSE, FALSE, FALSE, FALSE, TRUE];
    (* 逐台接管开关：TRUE = 该编号走真实硬件，FALSE = 走仿真。默认 1/2/3/6/8/9/10/17 为 TRUE。
    每次上电或完整下载都会回到这个组合；要临时关某一台，在线改位即可，但重启后恢复。
    索引对照（与 GVL_DeviceIds 的对照表完全一致，换算规则：D 编号=索引，G 编号+8=索引）：
      1=D1 送料皮带    2=D2 切割走刀    3=D3 盘刀旋转    4=D4 定长平移
      5=D5 定长升降    6=D6 定长光电    7=D7 机械手平移   8=D8 平台旋转
      9=G1 下压       10=G2 侧挡升降   11=G3 侧推       12=G4 流利条升降
      13=G5 喷油      14=G6 吹气       15=G7 机械手升降  16=G8 机械手夹爪
      17=G9 盘刀升降
    本版本只有 1、2、3、8（真实轴）、6（真实光电）与 9、10、11、17（真实气缸）已实现适配；
    其中 9（G1 下压）是左右双压板，共 4 个限位、2 路阀，设备索引仍按 1 个计；
    10（G2 侧挡）是 300/450/600 三缸一组，共 6 个限位、3 路阀，索引同样按 1 个计。
    其余编号置 TRUE 会立即报 3002，不会被静默当仿真跑。
    改本数组会让整机强制回 Stopped 并要求重新初始化，见 FB_Machine 的 wRealMask 变化检测。 *)
xRelativeVerify : BOOL; (* 相对验证模式：未回零的真实轴把 Position 解释为正向 d 再反向 d 的往返；回零成功后自动改走绝对定位。 *)
xInterlockBypass : BOOL; (* 预留：手动模式已默认不做机构互锁，本开关当前不影响判定；后续手动按需补互锁时再用。 *)
xSafetyBypass : BOOL; (* 安全许可旁路一级开关；默认 FALSE，必须与二级同时置位才生效。 *)
xSafetyBypassConfirm : BOOL; (* 安全许可旁路二级确认；默认 FALSE，防止误点单开关就旁路。 *)
xUseRealMaterial : BOOL := TRUE; (* TRUE 使用真实定长光电（设备 6）的到位信号；FALSE 继续由 FB_SimPlant 产生来料。 *)
lrVerifyDistance : LREAL := 1.0; (* 相对验证单段距离，mm；首轮建议 0.5~2.0，代码内再限幅 20。 *)
lrVerifyVelocity : LREAL := 2.0; (* 相对验证速度，mm/s；只用于未回零时的低速往返验证，不再兼作手动限速。 *)
lrVerifyAcceleration : LREAL := 50.0; (* 相对验证加速度，mm/s2。 *)
lrVerifyDeceleration : LREAL := 50.0; (* 相对验证减速度，mm/s2。 *)
tVerifyDwell : TIME := T#500MS; (* 正向到位后的停留，保证 Execute 拉低至少一个扫描以形成新上升沿。 *)
lrVerifyMeasuredByHand : LREAL; (* 人工用百分表量到的正向段实际位移，mm；用于核对轴单位标定。 *)
lrHomePosition : LREAL := 0.0; (* 预留：回零完成后的坐标由轴配置的“回零坐标”决定，MC_Homing 没有 Position 入口，本字段当前不参与下发。 *)
tHomeTimeout : TIME := T#30S; (* 单轴回零超时；超时报 2004，防止找不到原点时无限等待。 *)
lrManualVelocityMax : LREAL := 200.0; (* 手动模式速度上限，mm/s（旋转轴为每秒角度）；放在结构体末尾，避免新增字段让已有在线变量错位。 *)
END_STRUCT
END_TYPE

// Device/Application/00_Types/ST_MachineStatus
(* 模块说明：提供给监控和上位机的整机状态。可从主步骤、支线步骤、报警和互锁阻挡编号定位等待原因。 *)
TYPE ST_MachineStatus :
STRUCT
	eState : E_MachineState; (* 整机状态，见 E_MachineState；调试时先确认是否已初始化及处于正确模式。 *)
	eMode : E_MachineMode; (* 本地模式旋钮的当前选择：Manual 手动，Automatic 自动；上位机仅可读取。 *)
	eAutoStep : E_AutoStep; (* 自动主流程步骤；送料、避让、切割、收尾等状态见 E_AutoStep。 *)
	xSimulation : BOOL; (* TRUE 使用内部仿真；当前 FALSE 报未实现 3001，不会接管真实运动。 *)
	xRealBackendAvailable : BOOL; (* 真实设备适配是否已具备；当前框架固定 FALSE。 *)
	xRemoteStartStopAllowed : BOOL; (* 当前是否允许上位机启停，供只读状态发布；与物理手动/自动模式独立。 *)
	xInitialized : BOOL; (* 初始化完成标志；停止、运行中切换模式或故障会清除。 *)
	xReady : BOOL; (* 整机已经初始化并处于 Ready 状态，可接受自动启动；手动状态下不置该位。 *)
	xMaterialAtLength : BOOL; (* 定长光电到位状态；自动送料须先离开再到位，并满足 D5 下降。 *)
	xCycleComplete : BOOL; (* 一个扫描周期的整循环完成脉冲，可用于计数或上位机提示。 *)
	udiCycleCount : UDINT; (* 已完成的自动整循环计数；包括机械手移料等三路收尾。 *)
	udiAlarm : UDINT; (* 整机锁存报警码；0 无报警，1001 安全许可，3001 实机未接入，10000+索引为设备故障。 *)
	uiBlockedDevice : UINT; (* 本扫描最后一个被互锁阻挡的设备索引；0 表示无阻挡，可结合设备状态排查。 *)
	uiManualReject : UINT; (* 本扫描最后一个被拒绝的手动设备索引；0 无拒绝，检查相反按钮或动作类型。 *)
	uiClearLengthStep : UINT; (* 避让支线 P 的当前步骤：10 升起 D5，20 移开 D4，1000 完成。 *)
	uiClearTransferStep : UINT; (* 避让支线 Q 当前步骤：10 降 G4，20 松 G3，30 降 G2，1000 完成。 *)
	uiPostStep : UINT; (* 收尾总步骤：10 抬刀，20 抬压，30 等待三路完成，1000 结束。 *)
	uiReturnKnifeStep : UINT; (* 收尾支线 A：10 喷油，20 D2 回刀，1000 完成。 *)
	uiUnloadStep : UINT; (* 机械手移料支线 B 步骤，10..110 每步加 10，1000 完成；详见 FB_Unload。 *)
	uiResetLengthStep : UINT; (* 收尾支线 C：10 D4 定位，20 D5 下降，30 确认下降，1000 完成。 *)
	uiInitializeStep : UINT; (* 初始化步骤：10 整理刀/压/夹爪，20 避让，25 真实轴回零，30 初始定位，40 定长下降，1000 完成。 *)
	uiActiveMaterialModel : UINT; (* 已采纳的运行料型，取自运行配方；可能与尚未生效的参数区不同。 *)
	wRemoteAckSequence : WORD; (* 整机已处理的上位机命令序号；应结合 uiRemoteResult 判断是否接受。 *)
	uiRemoteResult : UINT; (* 远程处理结果：0 接受，1 未授权，2 不支持命令，3 状态/本地停止不允许，4 验证模式禁止自动，5 配方不合法。 *)
	xAnyRealDevice : BOOL; (* 是否有任意设备由真实轴接管；TRUE 时安全源与状态发布走混跑逻辑。 *)
	xRelativeVerify : BOOL; (* 当前是否处于相对验证模式；此模式下绝对位置不作生产依据，禁止启动自动。 *)
	xSafetyBypassed : BOOL; (* 安全许可是否由两级软件旁路放行；仅调试期可为 TRUE。 *)
	uiSafetySource : UINT; (* 安全许可来源：0 仿真源，1 真实源，2 调试旁路。 *)
	wRealDeviceMask : WORD; (* 真实设备接管掩码，第 i 位置位表示设备 i 走真实轴；供上位机核对。 *)
	uiInitReject : UINT; (* 初始化被拒绝的原因：0 未拒绝；回零已并入初始化流程，当前无拒绝分支，字段预留。 *)
	xRealAxesHomed : BOOL; (* 所有已接管的真实轴都已完成回零；未接真实轴时为 TRUE。 *)
	xRunState : BOOL; (* 运行态锁存：按启动置 TRUE，按停止、安全许可丢失或进故障清 FALSE；没有它无法区分"锁存未解除"和"按钮没接"。 *)
END_STRUCT
END_TYPE

// Device/Application/00_Types/E_MachineMode
(* 模块说明：操作模式。手动与自动分别提出动作请求，共用设备执行和互锁。 *)
{attribute 'qualified_only'}
TYPE E_MachineMode :
(
    Manual := 0, (* 手动点动/单机构调试 *)
    Automatic := 1 (* 自动循环工序 *)
);
END_TYPE

// Device/Application/00_Types/ST_Recipe
(* 模块说明：加工配方。初始化和自动启动时校验并复制到运行配方，避免运行中参数变化影响当前工序。 *)
TYPE ST_Recipe :
STRUCT
uiMaterialModel : UINT := 300; (* 料型选择，仅支持 300/450/600，对应 G2 三个侧挡气缸；不是位移。 *)
lrCutHome : LREAL := 100.0; (* D2 切割起点，也是回刀终点；切割终点 = 该位置 + lrCutLength。 *)
lrCutLength : LREAL := 900.0; (* D2 本次切割行程；配合 lrCutHome=100 得到终点 1000。 *)
lrCutVelocity : LREAL := 200.0; (* D2 切割进给速度，mm/s；900mm 约 5 秒走完。 *)
lrReturnVelocity : LREAL := 100.0; (* D2 回刀速度，mm/s；回刀行程长，与切割速度分开设置。 *)
lrPositionVelocity : LREAL := 10.0; (* 其余定位动作的公共请求速度，当前为仿真示例。 *)
lrBeltVelocity : LREAL := 10.0; (* D1 皮带运行速度请求，当前未换算到实际驱动器单位。 *)
lrSpindleVelocity : LREAL := 50.0; (* D3 盘刀运行速度请求，mm/s；不是已标定的实际转速。自动切割默认 50。 *)
lrLengthPosition : LREAL := 100.0; (* D4 定长检测工作位置；到位后再令 D5 下降。 *)
lrLengthClear : LREAL := 0.0; (* D4 切割前避让位置；移动前须 D5 升起。 *)
lrRotateAngle : LREAL := 30; (* D8 平台旋转目标角度，示例范围为正负 360，实机角度单位待标定。 *)
lrGripperFront : LREAL := 100.0; (* D7 机械手前进取料位置。 *)
lrGripperPull : LREAL := 200.0; (* D7 夹紧后拉料目标位置。 *)
lrGripperBack : LREAL := 50.0; (* D7 松开后的抬升后退位置；到位后先下降，再最终回位。 *)
lrGripperHome : LREAL := 0.0; (* D7 机械手下降后最终回位的位置。 *)
tSpray : TIME := T#300MS; (* 收尾支线 A 的喷油保持时间；该步结束后撤销喷油请求。 *)
tStepTimeout : TIME := T#30S; (* 单动作步骤超时时间；正常送料等料阶段不套用此超时。 *)
tCutTimeout : TIME := T#30S; (* D2 切割步专用超时，独立于 tStepTimeout；加在结构体末尾，避免新增字段让已有在线变量错位。 *)
END_STRUCT
END_TYPE

// Device/Application/00_Types/ST_DeviceStatus
(* 模块说明：单个设备的执行反馈。收到命令与完成命令是两个状态，不能只看忙标志判断完成。 *)
TYPE ST_DeviceStatus :
STRUCT
xReady : BOOL; (* 设备已使能且无故障，允许接收命令；不表示动作已经完成。 *)
xBusy : BOOL; (* 当前动作正在执行，定位完成或停止后清除。 *)
xActive : BOOL; (* 连续运行已建立或点动正在进行；定位动作完成后不保持该标志。 *)
xError : BOOL; (* 本设备或本子流程发生故障；具体原因见对应错误码。 *)
udiErrorID : UDINT; (* 错误码；0 表示无错误，设备或流程发生异常时赋值。 *)
udiAcceptedID : UDINT; (* 设备已接收的命令序号，用于区别尚未接收与正在执行。 *)
udiCompletedID : UDINT; (* 设备已完成的命令序号；应与本次 udiID 匹配后再切换步骤。 *)
lrPosition : LREAL; (* 实际或仿真反馈位置；气缸 0/1 的方向见设备编号说明。 *)
xRealActive : BOOL; (* TRUE 表示该编号当前由真实执行后端接管，不是仿真模型；默认 FALSE。 *)
xHomed : BOOL; (* 真实轴本次上电后已完成回零；仿真设备恒为 FALSE。回零成功前绝对定位会被拒绝。 *)
END_STRUCT
END_TYPE

// Device/Application/00_Types/E_DeviceAction
(* 模块说明：统一设备动作类型。未请求或停止时取消动作；定位完成依据本次命令序号判断。 *)
{attribute 'qualified_only'}
TYPE E_DeviceAction :
(
    None := 0, (* 无动作请求，取消当前动作 *)
    Position := 1, (* 定位到指定目标，等待本次序号完成 *)
    Run := 2, (* 保持连续运行请求 *)
    Jog := 3, (* 保持点动，速度正负决定方向 *)
    Stop := 4, (* 取消动作，停止运行 *)
    Home := 5 (* 回零：按轴配置的回零方式寻找原点，完成后把轴坐标设为回零坐标 *)
);
END_TYPE

// Device/Application/00_Types/E_MachineState
(* 模块说明：整机运行状态。停止或报警复位后须重新初始化，启动命令不会跳过初始化。 *)
{attribute 'qualified_only'}
TYPE E_MachineState :
(
    Stopped := 0, (* 停止，须初始化 *)
    Initializing := 10, (* 初始化中 *)
    Ready := 20, (* 初始化完成，等待自动启动 *)
    Manual := 30, (* 手动控制中 *)
    Automatic := 40, (* 自动工序运行中，包含正常等料 *)
    Fault := 90 (* 报警锁存，清除原因后复位 *)
);
END_TYPE

// Device/Application/00_Types/ST_DeviceCommand
(* 模块说明：上层发给单个设备的请求。定位每次换新序号；连续运行和点动期间保持请求。 *)
TYPE ST_DeviceCommand :
STRUCT
eAction : E_DeviceAction; (* 动作类型：无请求、定位、连续运行、点动或停止，见 E_DeviceAction。 *)
udiID : UDINT; (* 本次命令序号，0 无效；发起新定位时换新序号。 *)
lrTarget : LREAL; (* 目标工程位置；气缸使用约定的 0/1 端点，连续运行和点动不使用该位置。 *)
lrVelocity : LREAL; (* 请求速度，单位随设备工程单位定义；尚未完成实机标定。 *)
END_STRUCT
END_TYPE

// Device/Application/00_Types/ST_OperatorCommand
(* 模块说明：由本地实体面板解码形成的整机命令。模式取自旋钮，初始化/启动/复位取按钮；运行态由 FB_Machine 锁存。 *)
TYPE ST_OperatorCommand :
STRUCT
eMode : E_MachineMode := E_MachineMode.Manual; (* 本地模式旋钮的当前选择：Manual 手动，Automatic 自动；上位机仅可读取。 *)
xInitialize : BOOL; (* 初始化请求，上升沿有效；只允许从停止且许可满足时进入。 *)
xStart : BOOL; (* 自动启动请求，上升沿有效；须先初始化到 Ready。 *)
xStop : BOOL; (* 停止事件，兼容保留：远程停止帧仍会写一个扫描；物理停止按钮走 xRunStop。 *)
xResetAlarm : BOOL; (* 报警复位请求，上升沿有效；原因清除后复位，不会自动重新启动。 *)
xContinuous : BOOL; (* TRUE 连续循环；FALSE 在当前完整循环结束后回到就绪。 *)
xRunStart : BOOL; (* 启动按钮标准化电平，按一下一次上升沿；FB_Machine 用它的上升沿置运行态。 *)
xRunStop : BOOL; (* 停止按钮标准化电平（常闭已取反），按一下一次上升沿；FB_Machine 用它的上升沿清运行态。 *)
END_STRUCT
END_TYPE

// Device/Application/00_Types/ST_DeviceConfig
(* 模块说明：设备类型、行程范围和仿真参数。当前工程单位与时间均为仿真示例，尚未完成实机标定。 *)
TYPE ST_DeviceConfig :
STRUCT
	eKind : E_DeviceKind; (* 设备类型，决定调用哪一种设备适配功能块。 *)
	lrInitialPosition : LREAL; (* 首次进入仿真时的初始位置，不是实机回原点结果。 *)
	lrMinPosition : LREAL := -1000.0; (* 示例软行程下限，单位随机构定义。 *)
	lrMaxPosition : LREAL := 1000.0; (* 示例软行程上限，单位随机构定义。 *)
	lrMaxVelocity : LREAL := 100.0; (* 允许请求的最大速度，用于仿真命令范围检查。 *)
	tSimAction : TIME := T#500MS; (* 仿真单次定位/建立运行状态所需时间，不代表实际机械动作时间。 *)
	lrMaxAcceleration : LREAL := 50.0; (* 真实轴加速度上限，mm/s2；仿真不使用该字段。 *)
	lrMaxDeceleration : LREAL := 50.0; (* 真实轴减速度上限，mm/s2；仿真不使用该字段。 *)
	xAbsoluteAllowed : BOOL := FALSE; (* 真实轴是否允许绝对定位；未回零时必须保持 FALSE。 *)
END_STRUCT
END_TYPE

// Device/Application/00_Types/ST_SimulationSettings
(* 模块说明：软件仿真输入和异常注入。设备索引为 1..17，与 GVL_DeviceIds 一致。 *)
TYPE ST_SimulationSettings :
STRUCT
xSafetyOK : BOOL := TRUE; (* 安全许可接口或仿真许可，TRUE 允许；不等同于安全级急停回路。 *)
xAutoMaterial : BOOL := TRUE; (* TRUE 由仿真模型自动产生到位；FALSE 使用人工料到位输入。 *)
xMaterialSensor : BOOL; (* 手动模拟的光电到位信号，仅在 xAutoMaterial=FALSE 时使用。 *)
tMaterialDelay : TIME := T#1S; (* 满足皮带运行及定长下降条件后，仿真来料的延时时间。 *)
axStall : ARRAY[1..17] OF BOOL; (* 设备卡住注入，索引 1..17；保持忙且不完成，用于观察等待/超时。 *)
axFault : ARRAY[1..17] OF BOOL; (* 设备故障注入，索引 1..17；先清除注入，再执行报警复位。 *)
END_STRUCT
END_TYPE

// Device/Application/00_Types/E_DeviceKind
(* 模块说明：设备适配类型，由设备管理器选择轴、电机、气缸或阀的执行入口。 *)
{attribute 'qualified_only'}
TYPE E_DeviceKind :
(
    Unused := 0, (* 保留，不调度 *)
    Axis := 1, (* 定位轴 *)
    Motor := 2, (* 连续电机 *)
    Cylinder := 3, (* 两端动作气缸 *)
    Valve := 4 (* 开关阀 *)
);
END_TYPE

// Device/Application/00_Types/ST_ManualCommand
(* 模块说明：手动按钮接口。点动和运行按住有效，定位使用上升沿；手动请求同样经过互锁。 *)
TYPE ST_ManualCommand :
STRUCT
xJogPositive : BOOL; (* 手动正向点动，按住有效，释放后取消；只支持定位轴。 *)
xJogNegative : BOOL; (* 手动反向点动，按住有效；与正向同时按下会被拒绝。 *)
xMove : BOOL; (* 手动定位按钮，上升沿锁存目标，动作保持到本次序号完成。 *)
xHome : BOOL; (* 手动回零按钮，上升沿触发一次，动作保持到本次回零完成；只支持真实轴 D2/D8，D3 盘刀为连续旋转主轴不回零。 *)
xRun : BOOL; (* 手动连续运行按钮，按住有效、松开停止，仅支持 D1/D3/G5/G6；D3 接真实轴后由驱动器带载运行。 *)
lrTarget : LREAL; (* 目标工程位置；气缸使用约定的 0/1 端点，连续运行和点动不使用该位置。 *)
lrVelocity : LREAL := 100.0; (* 请求速度，单位随设备工程单位定义；尚未完成实机标定。 *)
END_STRUCT
END_TYPE

// Device/Application/00_Types/E_AutoStep
(* 模块说明：自动主流程步骤。正常循环从送料等料开始，切割完成后执行三路收尾。 *)
{attribute 'qualified_only'}
TYPE E_AutoStep :
(
    Idle := 0, (* 主流程待机 *)
    FeedWait := 10, (* 正常送料等料，可长期等待 *)
    StopFeed := 20, (* 撤销皮带运行并等待停止 *)
    Push := 30, (* G3 推动气缸动作 *)
    Clearance := 40, (* 并行避让 P/Q，全完成后继续 *)
    Rotate := 50, (* D8 平台旋转到配方角度 *)
    PressDown := 60, (* G1 下压到位 *)
    KnifeDown := 70, (* G9 盘刀下降到位 *)
    SpindleOn := 80, (* D3 盘刀运行状态建立 *)
    Cutting := 90, (* D2 走刀和 G6 吹气，等待指定行程到位 *)
    StopCut := 100, (* 停止盘刀和吹气 *)
    PostCut := 110, (* 抬刀、抬压、并行三路收尾 *)
    Complete := 120, (* 整循环完成，连续模式回送料 *)
    Fault := 900 (* 自动流程错误，退出执行后复位 *)
);
END_TYPE

// Device/Application/00_Types/ST_RemoteCommand
(* 模块说明：上位机可选启停请求，不含模式、初始化、复位或连续选择字段。参数通过独立配方接口下发。 *)
TYPE ST_RemoteCommand :
STRUCT
xStart : BOOL; (* 自动启动请求，上升沿有效；须先初始化到 Ready。 *)
xStop : BOOL; (* 普通停止，TRUE 持续有效；取消动作并清除初始化，不能替代硬件急停。 *)
END_STRUCT
END_TYPE

// Device/Application/00_Types/ST_PanelInputs
(* 模块说明：实体旋钮与按钮的逻辑输入；映射层先处理常开/常闭和极性，不在此处指定物理地址。仿真使用相同格式。 *)
TYPE ST_PanelInputs :
STRUCT
xAutoMode : BOOL; (* 模式旋钮的标准化逻辑值：TRUE 自动，FALSE 手动；不是上位机设定值。 *)
xInitialize : BOOL; (* 初始化请求，上升沿有效；只允许从停止且许可满足时进入。 *)
xStart : BOOL; (* 自动启动请求，上升沿有效；须先初始化到 Ready。 *)
xStop : BOOL; (* 停止事件，兼容保留：远程停止帧仍会写一个扫描；物理停止按钮不走这里。 *)
xResetAlarm : BOOL; (* 报警复位请求，上升沿有效；原因清除后复位，不会自动重新启动。 *)
xRunStart : BOOL; (* 启动按钮原始电平，常开、按下为 TRUE；上升沿在 FB_Machine 内锁存运行态。 *)
xRunStop : BOOL; (* 停止按钮标准化电平：常闭触点已在本层取反，按下为 TRUE；上升沿清除运行态。 *)
END_STRUCT
END_TYPE

// Device/Application/01_Data/GVL_Parameters
(* 模块说明：仿真开关和待执行配方。参数生效时机见 ST_Recipe；关闭仿真当前报 3001，未接入真实设备。 *)
VAR_GLOBAL
    (* 以下默认值仅供软件仿真，不能直接作为已确认的生产参数。 *)
    xSimulation : BOOL := TRUE; (* TRUE 使用内部仿真；当前 FALSE 报未实现 3001，不会接管真实运动。 *)
    xContinuous : BOOL := FALSE; (* 本地工程配置的单循环/连续选择；上位机启停帧不修改此设置，默认单循环。 *)
    xAllowRemoteStartStop : BOOL := FALSE; (* 本地工程配置授权远程启停，默认 FALSE；不授予改模式、初始化或复位权限，也不映射给上位机写。 *)
    stRecipe : ST_Recipe; (* 待执行配方：初始化和自动启动时校验并取快照，运行中修改不会立即生效。 *)
    xUseRealPanel : BOOL := TRUE; (* TRUE 读物理面板按钮/旋钮；FALSE 读仿真面板。与 xSimulation 解耦，后者恒为 TRUE。 *)
END_VAR

// Device/Application/01_Data/GVL_IO_Physical
(* 模块说明：物理 I/O 符号层——传感器与电磁阀的唯一入口。
   本 GVL 刻意不带 AT %I* / AT %Q* 地址：通道由 InoProShop 的 I/O 映射页手工绑定，
   因此增减模块、调整 Local Bus 顺序都不会让符号与通道错位（地址由编译器重排，符号绑定不变）。

   极性约定（软件语义固定，与接线方式解耦）：
     DO  TRUE = 阀得电 = 设备动作（下压 / 伸出 / 下降）
     DI  TRUE = 该端到位
   若现场接线极性相反，只在本层取反，不改上层任何流程或互锁代码。

   当前分配建议（硬件工程师可调整，调整后同步改本注释即可）：
     DO  GL20_0032ETN  QB(I) bit0..bit4  -> G1左 / G1右 / G2-300 / G2-450 / G2-600
     DO  GL20_0032ETN  QB(I) bit5..bit6  -> G9 / 备用
     DO  指示灯另分配                    -> 绿灯 / 红灯
     DI  GL20_3200END  DI00..DI09        -> G1左(2) G2-300(2) G3(2) G9(2) G1右(2)
     DI  新增 4 点                       -> G2-450(2) G2-600(2)

   注意：G2 从单缸改成 300/450/600 三缸后，输出多占 2 点、输入多占 4 点。
   3200END 的 16 点 DI 原本已用 10 点，加 4 点后剩 2 点，仍然不够面板 8 点用，
   面板输入必须另加一块 DI 模块（这一点与改造前结论一致）。
   旧符号 xDoG2Valve / xDiG2Retract / xDiG2Extend 已停用，保留仅为避免已画好的
   映射页断开时报“符号不存在”，物理通道改绑到下方三个新阀与六个新限位符号。
*)
VAR_GLOBAL
    (* ===== 数字输出：GL20-0032ETN，单电控阀，高电平使能 ===== *)
    xDoG1ValveL : BOOL; (* G1 左压板阀：TRUE=下压，FALSE=抬起。建议 QB(I) bit0。 *)
    xDoG1ValveR : BOOL; (* G1 右压板阀：与左阀同命令同步动作。建议 QB(I) bit1。 *)
    xDoG2Valve300 : BOOL; (* G2 料型 300 侧挡阀：TRUE=该缸下降挡料，FALSE=提升。建议 QB(I) bit2。 *)
    xDoG2Valve450 : BOOL; (* G2 料型 450 侧挡阀：TRUE=该缸下降挡料，FALSE=提升。建议 QB(I) bit3。 *)
    xDoG2Valve600 : BOOL; (* G2 料型 600 侧挡阀：TRUE=该缸下降挡料，FALSE=提升。建议 QB(I) bit4。 *)
    xDoG3Valve : BOOL; (* G3 侧推阀：TRUE=侧推，FALSE=退回。建议 QB(I) bit5。 *)
    xDoG9Valve : BOOL; (* G9 盘刀升降阀：TRUE=下降进刀，FALSE=提升。建议 QB(I) bit6。 *)

    (* ===== 已停用：G2 原单缸阀。物理接线改绑 xDoG2Valve300/450/600，本符号保留不复用。 ===== *)
    xDoG2Valve : BOOL; (* 停用：G2 单缸阀旧符号，程序不再写入，保留仅为兼容已有映射页。 *)

    (* ===== 面板指示灯：两个纯输出，只有电平没有反馈 ===== *)
    xDoLampGreen : BOOL; (* 绿灯：手动/就绪常亮，自动循环运行中慢闪。 *)
    xDoLampRed : BOOL; (* 红灯：停机或故障时常亮。 *)

    (* ===== 数字输入：GL20-3200END，G1 双压板 4 点 + G3/G9 各 2 点 + G2 三缸 6 点 ===== *)
    (* G1 下压左压板 *)
    xDiG1LRetract : BOOL; (* 左缸抬起到位。建议 DI00。 *)
    xDiG1LExtend : BOOL; (* 左缸下压到位。建议 DI01。 *)

    (* G2 侧挡 300 缸 *)
    xDiG2_300Retract : BOOL; (* 300 缸提升到位。建议 DI02。 *)
    xDiG2_300Extend : BOOL; (* 300 缸下降到位。建议 DI03。 *)

    (* G3 侧推气缸 *)
    xDiG3Retract : BOOL; (* G3 退回到位。建议 DI04。 *)
    xDiG3Extend : BOOL; (* G3 伸出到位。建议 DI05。 *)

    (* G9 盘刀升降 *)
    xDiG9Retract : BOOL; (* G9 提升到位。建议 DI06。 *)
    xDiG9Extend : BOOL; (* G9 下降到位。建议 DI07。 *)

    (* G1 下压右压板：与左压板同属设备索引 9，两组传感器必须同时到位才算该端到位 *)
    xDiG1RRetract : BOOL; (* 右缸抬起到位。建议 DI08。 *)
    xDiG1RExtend : BOOL; (* 右缸下压到位。建议 DI09。 *)

    (* G2 侧挡 450 / 600 缸：新增 4 点，3200END 已无空位，需另加 DI 模块或换 32 点模块 *)
    xDiG2_450Retract : BOOL; (* 450 缸提升到位。 *)
    xDiG2_450Extend : BOOL; (* 450 缸下降到位。 *)
    xDiG2_600Retract : BOOL; (* 600 缸提升到位。 *)
    xDiG2_600Extend : BOOL; (* 600 缸下降到位。 *)

    (* ===== 已停用：G2 原单缸限位。改用上方三缸各自的六个限位符号。 ===== *)
    xDiG2Retract : BOOL; (* 停用：G2 单缸提升到位旧符号，程序不再读取。 *)
    xDiG2Extend : BOOL; (* 停用：G2 单缸下降到位旧符号，程序不再读取。 *)

    (* ===== 定长光电：D6，遮挡=有料。通道由映射页手工绑定，接哪个模块哪一位都行 ===== *)
    xDiMaterialLength : BOOL; (* 定长光电：TRUE=被遮挡=料已到位。建议接在还空着的 DI 上。 *)

    (* ===== 预留：喷油 / 吹气（本轮不接，占位避免后期改结构） ===== *)
    xDoG5Spray : BOOL; (* 喷油阀：TRUE=喷油。待分配。 *)
    xDoG6Air : BOOL; (* 吹气阀：TRUE=吹气。待分配。 *)

    (* ===== 测试控制面板输入：符号名固定，通道同样由映射页手工绑定 ===== *)
    (* 极性：除急停与停止外，均为常开触点，按下/到位为 TRUE。 *)
    xDiPanelAutoMode : BOOL; (* 自动/手动旋钮：TRUE=自动，FALSE=手动。 *)
    xDiPanelSafetyPermit : BOOL; (* 安全许可旋钮：TRUE=许可。 *)
    xDiEStop : BOOL; (* 急停自锁按钮，常开，按下=TRUE=不安全；断线读 FALSE 软件无法分辨，需外部安全回路。 *)
    xDiPanelRunStart : BOOL; (* 启动按钮，常开，按下=TRUE；上升沿把整机置为运行态。 *)
    xDiPanelRunStop : BOOL; (* 停止按钮，常闭：未按=TRUE，按下=FALSE；逻辑层取反后按上升沿处理。 *)
    xDiPanelStart : BOOL; (* start 按钮，常开，按下=TRUE；自动循环启动，须已初始化到 Ready。 *)
    xDiPanelInit : BOOL; (* 初始化按钮，常开，按下=TRUE。 *)
    xDiPanelReset : BOOL; (* 报警复位按钮，常开，按下=TRUE。 *)
END_VAR

// Device/Application/01_Data/GVL_Modbus
(* 模块说明：Modbus 收发缓冲区，索引从 0 开始，尚未绑定网络寄存器。实际地址和字序需另行配置。 *)
VAR_GLOBAL
    (* 仅预留收发缓冲区，尚未绑定工程中的 MODBUS_TCP 网络映射。 *)
    xEnable : BOOL; (* 启用 Modbus 缓冲区解析，默认 FALSE；不代表网络映射已经配置。 *)
    awRx : ARRAY[0..31] OF WORD; (* v2 接收字：0=版本2，1=序号，2=命令2启动/3停止；3/4 保留且必须为0，不接受模式写入。 *)
    awTx : ARRAY[0..127] OF WORD; (* 发布字缓冲区 0..127；包含确认、状态、报警、计数和位置，详见程序内索引注释。 *)
END_VAR

// Device/Application/01_Data/GVL_RealDevice
(* 模块说明：真实设备接管设置的唯一入口。默认全部 FALSE，整机行为与改造前完全一致。 *)
VAR_GLOBAL
	stSettings : ST_RealDeviceSettings; (* 接管开关、验证参数、旁路开关集中在此，便于 HMI 与调试统一读写。 *)
END_VAR

// Device/Application/01_Data/GVL_DeviceIds
(* 模块说明：设备数组索引常量。D1..D8 对应索引 1..8，D6 保留；G1..G9 对应索引 9..17。

   全机所有设备数组共用这同一套 17 个索引，任何一处写错都会串到别人身上，所以先记住两条换算规则：
     D 编号 直接等于索引           D1..D8  ->  1..8
     G 编号 + 8 = 索引             G1..G9  ->  9..17

   ===== 17 个设备索引对照表 =====
   索引  代号  设备名称            类型       真实适配   绑定对象
   1     D1    送料皮带/输送轴     Axis       已接       songliao   点动/连续运行
   2     D2    切割走刀/回刀轴     Axis       已接       qiege      -
   3     D3    盘刀旋转电机        Axis       已接       pandao     按线性模式配置
   4     D4    定长平移轴          Axis       仿真       -          尚未接管
   5     D5    定长升降            Axis       仿真       -          0=升起避让，1=下降检测
   6     D6    定长光电            Sensor     已接       xDiMaterialLength 只读；TRUE=有料，遮挡即到位
   7     D7    机械手平移          Axis       仿真       -
   8     D8    平台旋转轴          Axis       已接       xuanzhuan  台达 ASDA-B3-E
   9     G1    下压气缸            Cylinder   已接       xDoG1ValveL/R  0=抬起，1=下压；左右双缸同动
   10    G2    侧挡升降（三缸）    Cylinder   已接       xDoG2Valve300/450/600 0=三缸全提，300/450/600=对应缸下降
   11    G3    推动气缸            Cylinder   已接       xDoG3Valve 0=放开，1=侧推
   12    G4    流利条升降          Cylinder   仿真       -          初始在提升端
   13    G5    喷油阀              Valve      仿真       xDoG5Spray 预留，待分配输出点
   14    G6    吹气阀              Valve      仿真       xDoG6Air   预留，待分配输出点
   15    G7    机械手升降          Cylinder   仿真       -          0=下降，1=提升
   16    G8    机械手夹爪          Cylinder   仿真       -          0=打开，1=夹紧
   17    G9    盘刀升降            Cylinder   已接       xDoG9Valve 0=提升，1=下降进刀

   报警码换算：整机报警 = 10000 + 索引。
     例：10001 = D1 皮带、10009 = G1 下压、10010 = G2 侧挡、10017 = G9 下刀。
     注意 10001 不是「1 号报警」，而是设备 1；真正的设备故障先看 udiErrorID 的千位。
   已在 FB_DeviceManager 中实现真实适配的编号：1、2、3、8（真实轴）、6（真实光电）与 9、10、11、17（真实气缸）。
   其余编号把 stReal.axRealDevice[i] 置 TRUE 会立即报 3002，不会被静默当仿真跑。 *)

VAR_GLOBAL CONSTANT
    D1_Belt : UINT := 1; (* D1 送料皮带电机，设备数组索引 1。 *)
    D2_CutFeed : UINT := 2; (* D2 切割走刀/回刀轴，设备数组索引 2。 *)
    D3_Spindle : UINT := 3; (* D3 盘刀旋转电机，设备数组索引 3。 *)
    D4_LengthMove : UINT := 4; (* D4 定长平移轴，设备数组索引 4。 *)
    D5_LengthLift : UINT := 5; (* D5 定长升降，0 升起避让，1 下降检测，索引 5。 *)
    D6_LengthSensor : UINT := 6; (* D6 定长光电（只读传感器），TRUE=有料，索引 6。 *)
    D7_GripperMove : UINT := 7; (* D7 机械手平移，索引 7；索引 6 为保留设备 D6。 *)
    D8_Rotate : UINT := 8; (* D8 平台旋转轴，设备数组索引 8。 *)
    G1_Press : UINT := 9; (* G1 下压气缸，0 抬起，1 下压，索引 9。 *)
    G2_SideStop : UINT := 10; (* G2 侧挡升降（三缸一组），目标 0=全提，300/450/600=对应缸下降，索引 10。 *)    (* G2 三个侧挡缸的料型号：同时作为设备 10 的命令目标值（lrTarget）和料型配方值（uiMaterialModel）。
       三者是同一套编号，不要再单独定义一套；界面上显示 300/450/600 就是这三个位号。 *)
    G2_Band300 : UINT := 300; (* G2 料型 300 对应的侧挡缸号。 *)
    G2_Band450 : UINT := 450; (* G2 料型 450 对应的侧挡缸号。 *)
    G2_Band600 : UINT := 600; (* G2 料型 600 对应的侧挡缸号。 *)
    G3_Push : UINT := 11; (* G3 推动气缸，0 放开，1 侧推，索引 11。 *)
    G4_RollerLift : UINT := 12; (* G4 流利条升降，0 下降，1 提升，索引 12。 *)
    G5_Spray : UINT := 13; (* G5 喷油阀，连续运行请求表示打开，索引 13。 *)
    G6_Air : UINT := 14; (* G6 吹气阀，切割开始打开、切割结束关闭，索引 14。 *)
    G7_GripperLift : UINT := 15; (* G7 机械手升降，0 下降，1 提升，索引 15。 *)
    G8_GripperClamp : UINT := 16; (* G8 机械手夹爪，0 打开，1 夹紧，索引 16。 *)
    G9_KnifeLift : UINT := 17; (* G9 盘刀升降，0 提升，1 下降，索引 17。 *)
END_VAR

// Device/Application/GVL_Motion
(* 模块说明：旧单轴 Demo 的操作和监控变量。新切割机框架不使用这些变量；旧 Demo 当前未挂周期任务。 *)
VAR_GLOBAL
    (* 旧 Demo 操作命令：仅供单轴测试，新整机流程不使用。 *)
    xEnable     : BOOL; (* 旧 Demo 的 pandao 伺服使能请求，TRUE 上使能，FALSE 关闭。 *)
    xReset      : BOOL; (* 旧 Demo 轴故障复位请求，接 MC_Reset.Execute。 *)
    xStop       : BOOL; (* 旧 Demo 停止请求；停止完成后释放锁定，再决定是否重新启动。 *)
    xJogFwd     : BOOL; (* 历史正向点动入口，当前旧 Demo 正文未接入。 *)
    xJogRev     : BOOL; (* 历史反向点动入口，当前旧 Demo 正文未接入。 *)
    xMoveRel    : BOOL; (* 历史相对定位入口，当前旧 Demo 正文未接入。 *)
    xMoveAbs    : BOOL; (* 历史绝对定位入口，当前旧 Demo 正文未接入。 *)
    xStartCycle : BOOL; (* 旧 Demo 单次往返启动，上升沿有效；当前 Demo 未周期调用。 *)

    rRelDist    : LREAL := 100.0; (* 历史单次相对距离 mm，当前往返正文不采用该参数。 *)
    rTargetPos  : LREAL := 0.0; (* 历史绝对目标位置 mm，当前往返正文不采用该参数。 *)

    (* 旧 Demo 运动参数：实际采用及限幅见各参数同行说明。 *)
    rJogVel     : LREAL := 10.0; (* 历史点动速度 mm/s，当前往返正文不采用该参数。 *)
    rVel        : LREAL := 30.0; (* 旧 Demo 往返速度 mm/s，正文限幅为 1..10。 *)
    rAcc        : LREAL := 200.0; (* 旧 Demo 加速度 mm/s²，正文限幅为 10..200。 *)
    rDec        : LREAL := 200.0; (* 旧 Demo 减速度 mm/s²，正文限幅为 10..200。 *)
    rStroke     : LREAL := 100.0; (* 旧 Demo 请求的单程距离 mm，正文使用绝对值并限制最大 20。 *)
    tDwell      : TIME  := T#1S; (* 旧 Demo 每个行程端点停留时间。 *)

    (* 旧 Demo 运行反馈：仅在旧程序被调用时更新。 *)
    xPowered    : BOOL; (* MC_Power.Status，伺服已使能反馈。 *)
    xAxisReady  : BOOL; (* 旧 Demo 中由已使能、非忙、无错误组合得到的可用标志。 *)
    xBusy       : BOOL; (* 往返功能块或停止功能块正忙。 *)
    xDisabled   : BOOL; (* 旧 Demo 根据未使能得到的显示状态。 *)
    xStandStill : BOOL; (* 旧 Demo 根据已使能且非忙得到的显示状态，不是独立轴状态读取。 *)
    xStopping   : BOOL; (* 停止功能块正在执行。 *)
    xErrorStop  : BOOL; (* 旧 Demo 综合错误显示，与 xAxisError 同步。 *)
    xAxisError  : BOOL; (* 使能、往返、复位或停止功能块任一报错。 *)
    iAxisErrorID: DWORD; (* 历史错误码显示变量，当前正文未更新，需读取实际功能块 ErrorID。 *)
    rActPos     : LREAL; (* MC_ReadActualPosition 返回的 pandao 实际位置，单位 mm。 *)
    iState      : INT; (* 旧 Demo 当前 iCycle 步骤镜像，便于在线监控。 *)
END_VAR

// Device/Application/01_Data/GVL_Simulation
(* 模块说明：仿真调试入口。可模拟来料、动作卡住、设备故障和安全许可丢失。 *)
VAR_GLOBAL
    stSettings : ST_SimulationSettings; (* 软件仿真参数，含来料方式和异常注入。 *)
    stPanelInputs : ST_PanelInputs; (* 仿真旋钮/按钮输入；xAutoMode 选择模式，其余按钮按住/释放模拟物理信号。 *)
END_VAR

// Device/Application/01_Data/GVL_Interface
(* 模块说明：监控与调试接口。stPanel 每周期由面板解码覆盖，不是上位机命令入口；手动请求保留待物理按钮映射。 *)
VAR_GLOBAL
    stPanel : ST_OperatorCommand; (* 本地面板解码结果，只读观察；每周期覆盖，操作请使用实体或仿真面板输入。 *)
    aManual : ARRAY[1..17] OF ST_ManualCommand; (* 各设备手动请求，索引 1..17；进入手动后先释放所有按钮再允许动作。 *)
    stStatus : ST_MachineStatus; (* 本模块对外发布的状态；字段含义见其数据类型。 *)
    aDeviceStatus : ARRAY[1..17] OF ST_DeviceStatus; (* 设备管理器汇总反馈，索引 1..17；供工序判断及在线监控。 *)
END_VAR

// Device/Application/01_Data/GVL_IO
(* 模块说明：逻辑 I/O 预留接口，尚未绑定物理地址。数字输出数组当前每周期清零；G2 当前料型仅用于观察。 *)
VAR_GLOBAL
    (* 当前均为普通逻辑变量，没有 AT %Q / %I 物理地址绑定。 *)
    xSafetyOK : BOOL; (* 安全许可接口或仿真许可，TRUE 允许；不等同于安全级急停回路。 *)
    stPanelInputs : ST_PanelInputs; (* 实体面板的模式旋钮、初始化、启动、停止、复位逻辑信号；急停走独立安全许可。 *)
    xMaterialAtLength : BOOL; (* 真实光电到位预留输入，当前未映射物理输入，仿真时不采用此值。 *)
    axDigitalInputs : ARRAY[0..31] OF BOOL; (* 预留数字输入位，索引 0..31；当前未映射到真实输入。 *)
    axDigitalOutputs : ARRAY[0..31] OF BOOL; (* 预留数字输出位，索引 0..31；当前由 FB_IOMap 每周期清 FALSE。 *)
    uiG2BandActive : UINT; (* G2 当前实际下降的料型带号 300/450/600；0 表示三缸全部提升，供诊断观察。 *)
END_VAR

// Device/Application/PLC_PRG
(* 模块说明：周期入口：先解码实体面板，再解析通信、调度整机、发布反馈和映射逻辑输出，仅在 ETHERCAT1 调用一次。 *)
PROGRAM PLC_PRG
VAR
	fbPanel : FB_PanelInput; (* 实体/仿真面板解码实例，须先于通信和整机调度调用。 *)
	fbCommunication : FB_ModbusInterface; (* 通信命令解析和状态打包实例；打包的是上一扫描已发布的整机反馈。 *)
	fbMachine : FB_Machine; (* 整机调度实例，包含初始化、手动、自动、互锁、报警和设备管理。 *)
	fbIO : FB_IOMap; (* 逻辑 I/O 映射实例，当前只形成诊断需求，不驱动真实输出。 *)
	fbLamp : FB_Indicator; (* 面板两色指示灯逻辑实例；纯输出，不参与控制。 *)
	xSafetyBypassActive : BOOL; (* 安全许可两级旁路已生效；仅当一级开关与二级确认同时置位。 *)
END_VAR

(* 本程序只在 ETHERCAT1 中周期调用一次；内部功能块沿本调用链每扫描执行。 *)
(* 0. 面板物理点 -> 逻辑面板：常开/常闭等极性只在这层处理，接线接反改这里一行即可。
   用 xUseRealPanel 而不是 xSimulation 选来源，因为 xSimulation 必须恒为 TRUE（FALSE 整机报 3001），
   真实设备是靠 axRealDevice 逐台接管的，物理按钮与设备仿真必须能同时存在。 *)
IF GVL_Parameters.xUseRealPanel THEN
    GVL_IO.stPanelInputs.xAutoMode   := GVL_IO_Physical.xDiPanelAutoMode;
    GVL_IO.stPanelInputs.xInitialize := GVL_IO_Physical.xDiPanelInit;
    GVL_IO.stPanelInputs.xStart      := GVL_IO_Physical.xDiPanelStart;
    GVL_IO.stPanelInputs.xResetAlarm := GVL_IO_Physical.xDiPanelReset;
    GVL_IO.stPanelInputs.xRunStart   := GVL_IO_Physical.xDiPanelRunStart;
    (* 停止按钮是常闭触点：未按=TRUE、按下=FALSE。这里取反成"TRUE=按下"，
       物理下降沿在逻辑层变回上升沿，FB_Machine 只认一个沿，不用分两种按钮。 *)
    GVL_IO.stPanelInputs.xRunStop    := NOT GVL_IO_Physical.xDiPanelRunStop;
    (* 安全许可 = 旋钮在许可位 且 急停未按下。急停是常开触点，按下=TRUE=不安全。
       注意这是联锁逻辑，不是安全级回路；断线时读到 FALSE 会被当成"许可成立"。 *)
    GVL_IO.xSafetyOK := GVL_IO_Physical.xDiPanelSafetyPermit AND NOT GVL_IO_Physical.xDiEStop;
ELSE
    (* 仿真面板调试：许可沿用仿真设置，物理旋钮与急停不参与，否则没有面板时永远过不了许可。 *)
    GVL_IO.xSafetyOK := GVL_Simulation.stSettings.xSafetyOK;
END_IF
(* 先解码实体/仿真面板；模式旋钮为唯一模式来源，随后发布到只读监控接口。 *)
fbPanel(xSimulation:=GVL_Parameters.xSimulation,stReal:=GVL_IO.stPanelInputs,
    stSim:=GVL_Simulation.stPanelInputs,xContinuous:=GVL_Parameters.xContinuous,
    xUseRealPanel:=GVL_Parameters.xUseRealPanel);
GVL_Interface.stPanel:=fbPanel.stCommand;
(* 1. 解析上位机新命令并打包上一扫描状态，供本扫描整机处理。 *)
fbCommunication(xEnable:=GVL_Modbus.xEnable,stStatus:=GVL_Interface.stStatus,
    aStatus:=GVL_Interface.aDeviceStatus,awRx:=GVL_Modbus.awRx,awTx:=GVL_Modbus.awTx);
(* 2. 安全许可旁路：一级开关与二级确认同时置位才生效，单开关无效。
   旁路只替代安全许可旋钮，绝不能盖掉急停：急停按下时旁路同样失效。 *)
xSafetyBypassActive:=F_SafetyBypassActive(GVL_RealDevice.stSettings) AND NOT GVL_IO_Physical.xDiEStop;
(* 3. 整机选择操作来源，调度工序，通过互锁后统一调用设备。 *)
fbMachine(
	xSimulation:=GVL_Parameters.xSimulation,
	stPanel:=GVL_Interface.stPanel,
    stRemote:=fbCommunication.stCommand,
	xRemoteRequest:=fbCommunication.xRequest,
    xAllowRemoteStartStop:=GVL_Parameters.xAllowRemoteStartStop,
    wRemoteSequence:=fbCommunication.wRequestSequence,
	aManual:=GVL_Interface.aManual,
    stRecipe:=GVL_Parameters.stRecipe,
	stSim:=GVL_Simulation.stSettings,
    stReal:=GVL_RealDevice.stSettings,
	xSafetyBypassActive:=xSafetyBypassActive,
    xRealSafetyOK:=GVL_IO.xSafetyOK,
	xRealMaterial:=GVL_IO.xMaterialAtLength);
(* 4. 将整机反馈发布到监控接口，建议调试时从这里查看主步骤和支线步骤。 *)
GVL_Interface.stStatus:=fbMachine.stStatus;
GVL_Interface.aDeviceStatus:=fbMachine.aDeviceStatus;

(* 4.5 定长光电（设备 6）接管后，把它本扫描的到位状态发布成真实料信号。
    这里取的是刚算完的设备状态；FB_Machine 内部读的是上一扫描的同一个值，
    对送料这种等稳定信号的判断没有影响（扫描周期远小于去抖时间）。 *)
GVL_IO.xMaterialAtLength := fbMachine.aDeviceStatus[6].xActive;
(* 5. 形成逻辑输出并下沉到物理点；真实气缸阀电平在此写入 GVL_IO_Physical。 *)
fbIO(aCommand:=fbMachine.aSelectedCommand,
        aStatus:=fbMachine.aDeviceStatus,aValveOut:=fbMachine.aValveOut,aValveOutAux:=fbMachine.aValveOutAux,
        aG2Valve:=fbMachine.aG2Valve,uiG2Band:=fbMachine.uiG2Band,
    axOutputs:=GVL_IO.axDigitalOutputs);
(* 6. 面板指示灯：只读整机状态，不参与任何控制，放在最后算以保证与本扫描状态一致。 *)
fbLamp(xRunState:=fbMachine.stStatus.xRunState,eState:=fbMachine.stStatus.eState,
    eMode:=fbMachine.stStatus.eMode,udiAlarm:=fbMachine.stStatus.udiAlarm);
GVL_IO_Physical.xDoLampGreen:=fbLamp.xGreen;
GVL_IO_Physical.xDoLampRed:=fbLamp.xRed;

END_PROGRAM

// Device/Application/04_Machine/FB_Machine
(* 模块说明：整机调度中心：命令选择、模式和报警管理、初始化/手动/自动调度、统一互锁、设备执行及状态发布。 *)
FUNCTION_BLOCK FB_Machine
VAR_INPUT
	xSimulation : BOOL; (* TRUE 使用内部仿真；当前 FALSE 报未实现 3001，不会接管真实运动。 *)
	stPanel : ST_OperatorCommand; (* 本地实体面板解码结果；模式、初始化、复位始终以它为准。 *)
	stRemote : ST_RemoteCommand; (* 上位机可选的启停请求，不包含模式或初始化/复位字段。 *)
	xRemoteRequest : BOOL; (* 远程新命令有效脉冲；无新帧时仅保留模式与连续选择。 *)
	xAllowRemoteStartStop : BOOL; (* 本地工程配置授权远程启停，默认 FALSE；不授予改模式、初始化或复位权限，也不映射给上位机写。 *)
	wRemoteSequence : WORD; (* 本次远程新命令序号，整机处理后写入确认状态。 *)
	aManual : ARRAY[1..17] OF ST_ManualCommand; (* 各设备手动请求，索引 1..17；进入手动后先释放所有按钮再允许动作。 *)
	stRecipe : ST_Recipe; (* 待校验配方或上层传入的运行配方，字段含义见 ST_Recipe。 *)
	stSim : ST_SimulationSettings; (* 软件仿真设置；设备管理器按设备索引读取卡住与故障注入。 *)
	stReal : ST_RealDeviceSettings; (* 真实设备接管设置；逐台位决定哪些编号走真实轴。 *)
	xRealSafetyOK : BOOL; (* 真实安全许可预留接口；当前仿真模式使用 stSim.xSafetyOK。 *)
	xRealMaterial : BOOL; (* 真实定长光电预留输入；当前仿真模式由 FB_SimPlant 提供。 *)
	xSafetyBypassActive : BOOL; (* 安全许可两级旁路已生效；仅在 xAnyReal 为 TRUE 时参与取或。 *)
END_VAR
VAR_OUTPUT
	stStatus : ST_MachineStatus; (* 本模块对外发布的状态；字段含义见其数据类型。 *)
	aDeviceStatus : ARRAY[1..17] OF ST_DeviceStatus; (* 设备管理器汇总反馈，索引 1..17；供工序判断及在线监控。 *)
	aSelectedCommand : ARRAY[1..17] OF ST_DeviceCommand; (* 通过统一互锁后的最终设备请求，交设备管理器执行。 *)
	aValveOut : ARRAY[1..17] OF BOOL; (* 各设备阀电气电平，索引同设备号；供物理映射层下沉到真实输出点。 *)
	aValveOutAux : ARRAY[1..17] OF BOOL; (* 第二个执行器的阀电气电平，索引同设备号；当前只有 G1 双压板使用。 *)
	aG2Valve : ARRAY[1..3] OF BOOL; (* G2 三个侧挡阀电气电平 1=300，2=450，3=600；供物理映射层下沉。 *)
	uiG2Band : UINT; (* G2 当前实际下降的料型带号 300/450/600；0 表示三缸全部提升。 *)
END_VAR
VAR
	stCommand : ST_OperatorCommand; (* 本周期选择并合并后的整机命令；本地停止始终优先于远程。 *)
	stActiveRecipe : ST_Recipe; (* 本次初始化/自动启动时采纳的配方快照，运行中不直接跟随参数区变化。 *)
	aRequest : ARRAY[1..17] OF ST_DeviceCommand; (* 初始化/手动/自动产生的原始请求，每周期先清空，再交互锁筛选。 *)
	stEmpty : ST_DeviceCommand; (* 默认全零设备命令，每周期用它清空原始请求，未被重新提出的动作自动取消。 *)
	fbDevices : FB_DeviceManager; (* 统一设备管理器，每周期调用一次，汇总各设备反馈。 *)
	fbManual : FB_ManualControl; (* 手动请求转换功能块，须处于手动并已释放全部按钮才使能。 *)
	fbAuto : FB_AutoCycle; (* 自动主流程功能块，仅在整机 Automatic 状态运行。 *)
	fbInitialize : FB_Initialize; (* 初始化功能块，仅在整机 Initializing 状态执行。 *)
	fbInterlocks : FB_Interlocks; (* 所有模式共用的软件互锁，输出最终允许的请求。 *)
	fbPlant : FB_SimPlant; (* 仿真整机来料模型；当前流程读取其上一扫描的到位反馈。 *)
	fbAlarm : FB_AlarmManager; (* 整机首报警锁存功能块。 *)
	rtInitialize : R_TRIG; (* 初始化按钮上升沿检测。 *)
	rtStart : R_TRIG; (* 自动启动按钮上升沿检测。 *)
	rtReset : R_TRIG; (* 报警复位按钮上升沿检测。 *)
	rtRunStart : R_TRIG; (* 启动按钮上升沿：置运行态锁存。 *)
	rtRunStop : R_TRIG; (* 停止按钮上升沿：清运行态锁存（常闭触点在映射层已取反）。 *)
	xRunState : BOOL; (* 运行态锁存：按一下启动置 TRUE，按一下停止/安全丢失/进故障清 FALSE；全机唯一的"允许动作"判据。 *)
	udiCounter : UDINT; (* 全机共享的动作序号计数器，通过引用传递；由 F_NextID 分配，0 不使用。 *)
	udiFault : UDINT; (* 本扫描整理出的报警原因；设备错误使用 10000+设备索引。 *)
	xSafetyOK : BOOL; (* 安全许可接口或仿真许可，TRUE 允许；不等同于安全级急停回路。 *)
	xMaterial : BOOL; (* 当前实际采用的来料信号，仿真与实机预留输入二选一。 *)
	xInitialized : BOOL; (* 初始化完成标志；停止、运行中切换模式或故障会清除。 *)
	xPermit : BOOL; (* 整机当前允许发出动作的总许可；仍需继续满足各设备互锁。 *)
	xRemoteAccepted : BOOL; (* 本扫描远程命令已获授权，用于回传状态拒绝或配方错误。 *)
	xStartRequest : BOOL; (* 本次启动事件=本地启动按钮上升沿或已接受的远程启动帧；两种事件分别处理以免相互吞掉。 *)
	xResetDevices : BOOL; (* 本扫描设备复位脉冲，需复位上升沿、安全许可和仿真模式均满足。 *)
	xLastSimulation : BOOL := TRUE; (* 上扫描仿真开关；切换模式时清除初始化并停止。 *)
	xManualReleased : BOOL; (* 所有手动按钮都已释放，用于避免带着按住命令进入手动。 *)
	xManualArmed : BOOL; (* 本次进入手动后已观察到全部按钮释放；离开手动即清除。 *)
	eActiveMode : E_MachineMode; (* 当前初始化/运行时采纳的操作模式，用于检测运行中切换模式。 *)
	xAnyReal : BOOL; (* 是否有任意设备由真实轴接管；全 FALSE 时后续分支与改造前逐语句一致。 *)
    udiInterlockFault : UDINT; (* 互锁违规码；互锁在报警汇总之后才调用，故本扫描存入、下扫描并入 udiFault。 *)
	xAllHomed : BOOL; (* 所有已接管的真实轴都已完成回零；未接真实轴时为 TRUE，用于状态发布。 *)
	dwRealMask : DWORD; (* 真实设备接管掩码，第 i 位置位表示设备 i 走真实轴；用 DWORD 是因为索引 17 需要第 16 位，WORD 会溢出丢位。 *)
	dwLastRealMask : DWORD; (* 上扫描接管掩码；变化时清除初始化并回 Stopped。 *)
	xLastRelativeVerify : BOOL; (* 上扫描相对验证开关；切换时清除初始化并回 Stopped。 *)
	uiSafetySource : UINT; (* 安全许可来源：0 仿真源，1 真实源，2 调试旁路。 *)
	uiInitReject : UINT; (* 初始化被拒绝的原因：0 未拒绝；回零已并入初始化流程，当前无拒绝分支，字段预留。 *)
	i : INT; (* 本扫描数组遍历索引；含义及范围以当前 FOR 循环为准。 *)
END_VAR

(* 零、派生混跑标志：axRealDevice 全 FALSE 时 xAnyReal 为 FALSE，后续所有分支与改造前一致。 *)
xAnyReal:=FALSE; dwRealMask:=0;
FOR i:=1 TO 17 DO
    IF stReal.axRealDevice[i] THEN
        xAnyReal:=TRUE;
        dwRealMask:=dwRealMask OR SHL(DWORD#1,i-1);
    END_IF
END_FOR

(* 一、选择命令来源：本地默认优先；远程须授权，本地停止始终有效。 *)
stCommand:=stPanel;
(* 运行态锁存：按一下切换，不靠按钮保持。停止优先——同扫描两个都按下取停止。
   这是全机唯一的"允许动作"判据；下游不再出现单个按钮电平。 *)
rtRunStart(CLK:=stCommand.xRunStart);
rtRunStop(CLK:=stCommand.xRunStop);
IF rtRunStart.Q THEN xRunState:=TRUE; END_IF
IF rtRunStop.Q OR stCommand.xStop THEN xRunState:=FALSE; END_IF
(* 模式、初始化、复位来自实体面板；远程只可追加经过授权的启停，不能替换整份本地命令。 *)
xRemoteAccepted:=FALSE;
IF xRemoteRequest THEN
    stStatus.wRemoteAckSequence:=wRemoteSequence;
    IF xAllowRemoteStartStop THEN
        IF stRemote.xStop THEN
            stCommand.xStop:=TRUE;
            stStatus.uiRemoteResult:=0; xRemoteAccepted:=TRUE;
        ELSIF stRemote.xStart THEN
            IF (stPanel.eMode=E_MachineMode.Automatic)
               AND (stStatus.eState=E_MachineState.Ready) AND xRunState THEN
                stStatus.uiRemoteResult:=0; xRemoteAccepted:=TRUE;
            ELSE stStatus.uiRemoteResult:=3; END_IF
        ELSE stStatus.uiRemoteResult:=2; END_IF
    ELSE stStatus.uiRemoteResult:=1;
    END_IF
END_IF
(* 二、提取初始化/启动/复位上升沿；采样仿真或真实预留输入。 *)
rtInitialize(CLK:=stCommand.xInitialize);
rtStart(CLK:=stCommand.xStart);
(* 本地启动取按钮上升沿，远程启动取新帧脉冲，分别形成事件；本地停止仍优先。 *)
xStartRequest:=rtStart.Q OR (xRemoteAccepted AND stRemote.xStart AND NOT stRemote.xStop);
rtReset(CLK:=stCommand.xResetAlarm);
(* 混跑时安全源改为真实优先：未接安全回路时靠两级旁路放行，旁路生效不报 1001。 *)
IF xAnyReal THEN
    xSafetyOK:=xRealSafetyOK OR xSafetyBypassActive;
    IF stReal.xUseRealMaterial THEN xMaterial:=xRealMaterial;
    ELSE xMaterial:=fbPlant.xMaterialAtLength; END_IF
ELSIF xSimulation THEN xSafetyOK:=stSim.xSafetyOK; xMaterial:=fbPlant.xMaterialAtLength;
ELSE xSafetyOK:=xRealSafetyOK; xMaterial:=xRealMaterial; END_IF
(* 安全许可丢失立即清运行态：急停或旋钮离开许可位后，恢复必须重新按启动，不能自己回到运行。 *)
IF NOT xSafetyOK THEN xRunState:=FALSE; END_IF
(* 安全来源：0 仿真源，1 真实源，2 调试旁路。 *)
IF NOT xAnyReal THEN uiSafetySource:=0;
ELSIF xSafetyBypassActive AND NOT xRealSafetyOK THEN uiSafetySource:=2;
ELSE uiSafetySource:=1; END_IF
(* 三、整理当前报警原因并清空本扫描请求；未被子流程重新提出的动作自动取消。 *)
udiFault:=0;
IF NOT xSafetyOK THEN udiFault:=1001; END_IF
IF udiInterlockFault<>0 THEN udiFault:=udiInterlockFault; END_IF
IF NOT xSimulation THEN udiFault:=3001; END_IF
(* 仿真开关、接管掩码或验证模式变化，均清除初始化并回 Stopped。 *)
IF (xSimulation<>xLastSimulation) OR (dwRealMask<>dwLastRealMask) OR (stReal.xRelativeVerify<>xLastRelativeVerify) THEN
    stStatus.eState:=E_MachineState.Stopped; xInitialized:=FALSE;
END_IF
xLastSimulation:=xSimulation; dwLastRealMask:=dwRealMask; xLastRelativeVerify:=stReal.xRelativeVerify;
FOR i:=1 TO 17 DO
    IF aDeviceStatus[i].xError THEN udiFault:=10000+INT_TO_UDINT(i); END_IF
    aRequest[i]:=stEmpty;
END_FOR
(* 四、运行中切模式、停止或故障会撤销初始化，不能直接接续上一次工序。 *)
IF (stStatus.eState=E_MachineState.Automatic) OR (stStatus.eState=E_MachineState.Manual) THEN
    IF stCommand.eMode<>eActiveMode THEN stStatus.eState:=E_MachineState.Stopped; xInitialized:=FALSE; END_IF
END_IF
(* 停止是运行态锁存的电平判据：按一下停止后锁存一直为 FALSE，直到再按启动。
   这里用 xRunState 而不是按钮电平，是为了让"停着"和"按钮松开"不再有区别。 *)
IF NOT xRunState THEN
    IF (stStatus.eState<>E_MachineState.Stopped) AND (stStatus.eState<>E_MachineState.Fault) THEN
        stStatus.eState:=E_MachineState.Stopped;
    END_IF
    xInitialized:=FALSE;
END_IF
IF udiFault<>0 THEN stStatus.eState:=E_MachineState.Fault; xInitialized:=FALSE; END_IF
(* 五、复位设备和首报警锁存；必须先撤销故障原因，复位不自动启动。 *)
xResetDevices:=rtReset.Q AND xSafetyOK AND xSimulation;
IF xResetDevices THEN
    (* 复位时先按仍有效的故障注入判断原因，再清设备错误和整机锁存；原因未撤销不能复位。 *)
    udiFault:=0;
    udiInterlockFault:=0;
    FOR i:=1 TO 17 DO IF stSim.axFault[i] THEN udiFault:=10000+INT_TO_UDINT(i); END_IF END_FOR
END_IF
fbAlarm(udiIncoming:=udiFault,xReset:=xResetDevices);
IF (stStatus.eState=E_MachineState.Fault) AND (fbAlarm.udiLatched=0) AND xResetDevices THEN
    stStatus.eState:=E_MachineState.Stopped;
END_IF
IF fbAlarm.udiLatched<>0 THEN stStatus.eState:=E_MachineState.Fault; END_IF
(* 六、仅停止态接受初始化；配方通过检查后取快照。 *)
IF rtInitialize.Q AND xRunState THEN
    (* 真实轴的回零已并入初始化第 25 步，这里不再要求预先打开相对验证。 *)
    IF (stStatus.eState=E_MachineState.Stopped) AND xSimulation AND xSafetyOK AND F_RecipeValid(stRecipe) THEN
        stActiveRecipe:=stRecipe; stStatus.eState:=E_MachineState.Initializing;
        eActiveMode:=stCommand.eMode; xInitialized:=FALSE; uiInitReject:=0;
    ELSE
        (* 当前无拒绝分支：回零并入初始化，uiInitReject 保留字段但不再置位。 *)
        IF xRemoteAccepted THEN stStatus.uiRemoteResult:=3; END_IF
    END_IF
END_IF
(* 七、手动不依赖初始化：停机态只要模式在手动且运行态成立就直接进入，开机后不必先跑初始化。
   自动仍必须先完成初始化到 Ready；按过停止后运行态为假，手动也进不去，必须重新按启动。 *)
IF (stStatus.eState=E_MachineState.Stopped) AND (stCommand.eMode=E_MachineMode.Manual)
   AND xRunState THEN
    stStatus.eState:=E_MachineState.Manual; eActiveMode:=E_MachineMode.Manual;
END_IF
IF stStatus.eState=E_MachineState.Ready THEN
    IF stCommand.eMode=E_MachineMode.Manual THEN
        stStatus.eState:=E_MachineState.Manual; eActiveMode:=E_MachineMode.Manual;
    ELSIF xStartRequest AND xRunState THEN
        IF stReal.xRelativeVerify THEN
            (* 相对验证模式下绝对位置不作生产依据，禁止进自动。 *)
            stStatus.uiRemoteResult:=4;
        ELSIF F_RecipeValid(stRecipe) THEN
            stActiveRecipe:=stRecipe; eActiveMode:=E_MachineMode.Automatic;
            stStatus.eState:=E_MachineState.Automatic;
        ELSIF xRemoteAccepted THEN stStatus.uiRemoteResult:=5;
        END_IF
    END_IF
ELSIF (stStatus.eState=E_MachineState.Manual) AND (stCommand.eMode=E_MachineMode.Automatic) THEN
    stStatus.eState:=E_MachineState.Stopped; xInitialized:=FALSE;
END_IF
IF xStartRequest AND xRemoteAccepted AND (stStatus.eState<>E_MachineState.Automatic)
   AND (stStatus.uiRemoteResult=0) THEN stStatus.uiRemoteResult:=3; END_IF

(* 八、手动进入联锁：观察到一次全部按钮释放后，才开放点动/定位操作。 *)
xManualReleased:=TRUE;
FOR i:=1 TO 17 DO
    IF aManual[i].xJogPositive OR aManual[i].xJogNegative OR aManual[i].xMove OR aManual[i].xRun OR aManual[i].xHome THEN xManualReleased:=FALSE; END_IF
END_FOR
IF stStatus.eState<>E_MachineState.Manual THEN xManualArmed:=FALSE;
ELSIF xManualReleased THEN xManualArmed:=TRUE;
END_IF
(* 九、每扫描调用各模式功能块，失能的流程同时复位；共享请求只由当前模式提出。 *)
fbInitialize(xExecute:=stStatus.eState=E_MachineState.Initializing,stRecipe:=stActiveRecipe,
    aCommand:=aRequest,aStatus:=aDeviceStatus,udiCounter:=udiCounter);
fbManual(xEnable:=(stStatus.eState=E_MachineState.Manual) AND xManualArmed,stReal:=stReal,
    aManual:=aManual,aCommand:=aRequest,aStatus:=aDeviceStatus,udiCounter:=udiCounter);
fbAuto(xRun:=stStatus.eState=E_MachineState.Automatic,xContinuous:=stCommand.xContinuous,
    xMaterialAtLength:=xMaterial,stRecipe:=stActiveRecipe,aCommand:=aRequest,aStatus:=aDeviceStatus,udiCounter:=udiCounter);
(* 十、汇总流程完成和流程错误，单循环完成后回到 Ready。 *)
IF fbInitialize.xDone THEN xInitialized:=TRUE; stStatus.eState:=E_MachineState.Ready; END_IF
IF fbInitialize.xError OR fbAuto.xError THEN
    udiFault:=MAX(fbInitialize.udiErrorID,fbAuto.udiErrorID);
    fbAlarm(udiIncoming:=udiFault,xReset:=FALSE);
    stStatus.eState:=E_MachineState.Fault; xInitialized:=FALSE;
END_IF
IF fbAuto.xDone THEN
    stStatus.udiCycleCount:=stStatus.udiCycleCount+1;
    IF NOT stCommand.xContinuous THEN stStatus.eState:=E_MachineState.Ready; END_IF
END_IF
(* 十一、总许可与机构互锁筛选请求，再调用设备管理器；流程判断使用此前的反馈。 *)
xPermit:=xSimulation AND xSafetyOK AND xRunState AND (fbAlarm.udiLatched=0)
    AND ((stStatus.eState=E_MachineState.Initializing) OR (stStatus.eState=E_MachineState.Manual)
    OR (stStatus.eState=E_MachineState.Automatic));
(* 互锁违规先清后置：违规在下面 fbInterlocks 之后才算出，本扫描存入，下扫描并入 udiFault。 *)
udiInterlockFault:=0;
fbInterlocks(xPermit:=xPermit,xManualMode:=(stStatus.eState=E_MachineState.Manual),
    stRecipe:=stActiveRecipe,stReal:=stReal,aRequest:=aRequest,aStatus:=aDeviceStatus);
aSelectedCommand:=fbInterlocks.aCommand;
IF fbInterlocks.xViolated THEN udiInterlockFault:=5000+UINT_TO_UDINT(fbInterlocks.uiViolatedDevice); END_IF
fbDevices(xEnable:=xSimulation AND xSafetyOK,xSimulation:=xSimulation,xReset:=xResetDevices,
    xFaultHold:=(fbAlarm.udiLatched<>0),stSim:=stSim,stReal:=stReal,
    uiMaterialModel:=stActiveRecipe.uiMaterialModel,aCommand:=aSelectedCommand);
aDeviceStatus:=fbDevices.aStatus;
aValveOut:=fbDevices.aValveOut;
aValveOutAux:=fbDevices.aValveOutAux;
aG2Valve:=fbDevices.aG2Valve;
uiG2Band:=fbDevices.uiG2Band;
fbPlant(xEnable:=xSimulation,stSettings:=stSim,aStatus:=aDeviceStatus);
(* 十二、集中发布状态；机械手/定长/回刀卡在哪一步，可从对应 ui...Step 追踪。 *)
(* 故障一律清运行态：故障原因消失后不会自己恢复运行，必须重新按启动。 *)
IF stStatus.eState=E_MachineState.Fault THEN xRunState:=FALSE; END_IF
stStatus.eMode:=stCommand.eMode; stStatus.eAutoStep:=fbAuto.eStep;
stStatus.xSimulation:=xSimulation; stStatus.xRealBackendAvailable:=xAnyReal;
(* 对外掩码仍是 WORD，索引 17（第 16 位）不进这个字段；看真实接管请用 dwRealMask 内部量。 *)
stStatus.xAnyRealDevice:=xAnyReal; stStatus.wRealDeviceMask:=DWORD_TO_WORD(dwRealMask);
stStatus.xRunState:=xRunState;
stStatus.xRelativeVerify:=stReal.xRelativeVerify;
stStatus.xSafetyBypassed:=xSafetyBypassActive AND xAnyReal;
stStatus.uiSafetySource:=uiSafetySource; stStatus.uiInitReject:=uiInitReject;
stStatus.xRemoteStartStopAllowed:=xAllowRemoteStartStop;
xAllHomed:=TRUE;
FOR i:=1 TO 17 DO
    (* D3 盘刀只做连续旋转、不做回零，不参与“全部真实轴已回零”判定，否则该状态永远为 FALSE。 *)
    IF stReal.axRealDevice[i] AND (i<>3) AND (i<9) AND NOT aDeviceStatus[i].xHomed THEN xAllHomed:=FALSE; END_IF
END_FOR
stStatus.xRealAxesHomed:=xAllHomed;
stStatus.xInitialized:=xInitialized;
stStatus.xReady:=xInitialized AND (stStatus.eState=E_MachineState.Ready);
stStatus.xMaterialAtLength:=xMaterial; stStatus.xCycleComplete:=fbAuto.xDone;
stStatus.udiAlarm:=fbAlarm.udiLatched; stStatus.uiBlockedDevice:=fbInterlocks.uiBlockedDevice;
stStatus.uiManualReject:=fbManual.uiRejectDevice;
stStatus.uiClearLengthStep:=fbAuto.uiClearLengthStep; stStatus.uiClearTransferStep:=fbAuto.uiClearTransferStep;
stStatus.uiPostStep:=fbAuto.uiPostStep; stStatus.uiReturnKnifeStep:=fbAuto.uiReturnKnifeStep;
stStatus.uiUnloadStep:=fbAuto.uiUnloadStep; stStatus.uiResetLengthStep:=fbAuto.uiResetLengthStep;
stStatus.uiInitializeStep:=fbInitialize.uiStep; stStatus.uiActiveMaterialModel:=stActiveRecipe.uiMaterialModel;

END_FUNCTION_BLOCK

// Device/Application/04_Machine/F_RecipeValid
(* 模块说明：检查框架允许的料型、速度、行程和位置顺序。通过仅表示符合示例边界，不代表实机参数已经确认。 *)
FUNCTION F_RecipeValid : BOOL
VAR_INPUT
    stRecipe : ST_Recipe; (* 待校验配方或上层传入的运行配方，字段含义见 ST_Recipe。 *)
END_VAR

(* 示例边界：切长 0..1200、速度 0..300、角度正负360，并要求机械手回位<后退<前进<拉料。边界是否适合实机仍需标定。 *)
(* 料型只认 300/450/600：现场侧挡是三个固定位置的气缸，没有 400 这个档；400 是早期仿真的占位值。 *)
F_RecipeValid := ((stRecipe.uiMaterialModel = 300) OR
    (stRecipe.uiMaterialModel = 450) OR (stRecipe.uiMaterialModel = 600))
    AND (stRecipe.lrCutLength > 0.0) AND (stRecipe.lrCutLength <= 1200.0)
    AND (stRecipe.lrCutVelocity > 0.0) AND (stRecipe.lrCutVelocity <= 300.0)
    AND (stRecipe.lrReturnVelocity > 0.0) AND (stRecipe.lrReturnVelocity <= 300.0)
    AND (stRecipe.lrPositionVelocity > 0.0) AND (stRecipe.lrPositionVelocity <= 100.0)
    AND (stRecipe.lrBeltVelocity > 0.0) AND (stRecipe.lrBeltVelocity <= 100.0)
    AND (stRecipe.lrSpindleVelocity > 0.0) AND (stRecipe.lrSpindleVelocity <= 100.0)
    AND (stRecipe.tStepTimeout >= T#1S) AND (stRecipe.tCutTimeout >= T#1S) AND (stRecipe.tSpray > T#0MS)
    AND (ABS(stRecipe.lrCutHome) <= 500.0)
    (* 终点 = 回刀起点 + 切割行程；行程放到 1200 后，终点上限相应放到 1300（典型 100+1200）。 *)
    AND (ABS(stRecipe.lrCutHome + stRecipe.lrCutLength) <= 1300.0)
    AND (ABS(stRecipe.lrLengthPosition) <= 1000.0)
    AND (ABS(stRecipe.lrLengthClear) <= 1000.0)
    AND (ABS(stRecipe.lrRotateAngle) <= 360.0)
    AND (stRecipe.lrGripperHome < stRecipe.lrGripperBack)
    AND (stRecipe.lrGripperBack < stRecipe.lrGripperFront)
    AND (stRecipe.lrGripperFront < stRecipe.lrGripperPull)
    AND (ABS(stRecipe.lrGripperPull) <= 1000.0);

END_FUNCTION

// Device/Application/06_Simulation/FB_SimPlant
(* 模块说明：仿真来料模型。皮带运行且定长下降时延时产生一次到位，定长升起或关闭模型后清除。 *)
FUNCTION_BLOCK FB_SimPlant
VAR_INPUT
    xEnable : BOOL; (* 本功能使能，电平有效；失能时不接受新的动作请求。 *)
    stSettings : ST_SimulationSettings; (* 软件仿真参数，含来料方式和异常注入。 *)
    aStatus : ARRAY[1..17] OF ST_DeviceStatus; (* 各设备的反馈数组 1..17，供判断忙、完成序号、故障和位置。 *)
END_VAR
VAR_OUTPUT
    xMaterialAtLength : BOOL; (* 定长光电到位状态；自动送料须先离开再到位，并满足 D5 下降。 *)
END_VAR
VAR
    xLatched : BOOL; (* 本轮仿真料到位保持标志；定长升起或模型失能时清除。 *)
    tonMaterial : TON; (* 自动仿真来料延时，仅在运行皮带且定长下降到位时计时。 *)
END_VAR

(* 定长抬起时清除上次来料；自动方式形成一次延时到位，手动方式直接采用人工传感器。 *)
IF NOT xEnable OR NOT F_At(aStatus[5],1.0) THEN xLatched:=FALSE; END_IF
tonMaterial(IN:=xEnable AND stSettings.xAutoMaterial AND aStatus[1].xActive
    AND F_At(aStatus[5],1.0) AND NOT xLatched,PT:=stSettings.tMaterialDelay);
IF tonMaterial.Q THEN xLatched:=TRUE; END_IF
IF stSettings.xAutoMaterial THEN xMaterialAtLength:=xLatched;
ELSE xMaterialAtLength:=xEnable AND F_At(aStatus[5],1.0) AND stSettings.xMaterialSensor;
END_IF

END_FUNCTION_BLOCK

// Device/Application/02_Devices/F_At
(* 模块说明：检查设备可用、无忙无故障且位置误差小于 0.01。它检查位置，不检查本次命令序号。 *)
FUNCTION F_At : BOOL
VAR_INPUT
    stStatus : ST_DeviceStatus; (* 本模块对外发布的状态；字段含义见其数据类型。 *)
    lrTarget : LREAL; (* 要检查的目标位置；误差小于 0.01 且设备就绪、无忙无错时返回 TRUE。 *)
END_VAR

(* 位置容差为 0.01 工程单位；这里不做新命令序号校验，用于姿态/互锁判断。 *)
F_At := stStatus.xReady AND NOT stStatus.xBusy
    AND NOT stStatus.xError AND (ABS(stStatus.lrPosition-lrTarget) < 0.01);

END_FUNCTION

// Device/Application/02_Devices/FB_DeviceManager
FUNCTION_BLOCK FB_DeviceManager
(* 模块说明：统一设备执行入口。首次建立类型和初始位置，每扫描周期按类型调用设备功能块并收集反馈。 *)
VAR_INPUT
	xEnable : BOOL; (* 本功能使能，电平有效；失能时不接受新的动作请求。 *)
	xSimulation : BOOL; (* TRUE 使用内部仿真；当前 FALSE 报未实现 3001，不会接管真实运动。 *)
	xReset : BOOL; (* 故障复位许可；仿真设备仅在故障注入已撤销时清除错误。 *)
	xFaultHold : BOOL; (* 整机故障保持：TRUE 时真实轴强制停车、真实阀失电，直到复位。 *)
	stSim : ST_SimulationSettings; (* 软件仿真设置；设备管理器按设备索引读取卡住与故障注入。 *)
	stReal : ST_RealDeviceSettings; (* 真实设备接管设置；逐台位决定该编号走真实轴还是仿真。 *)
	uiMaterialModel : UINT; (* 当前运行料型 300/450/600；G2 气缸组按此选通其中一个缸下降。 *)
	aCommand : ARRAY[1..17] OF ST_DeviceCommand; (* 统一设备请求数组 1..17；子流程写请求，设备管理器执行。 *)
END_VAR
VAR_OUTPUT
	aStatus : ARRAY[1..17] OF ST_DeviceStatus; (* 各设备的反馈数组 1..17，供判断忙、完成序号、故障和位置。 *)
	aValveOut : ARRAY[1..17] OF BOOL; (* 各设备的阀电气输出电平 1..17；只有已接管的真实气缸可能为 TRUE，供物理映射层取用。 *)
	aValveOutAux : ARRAY[1..17] OF BOOL; (* 第二个执行器的阀电气电平 1..17；当前只有 G1 双压板的 [9] 有效，其余恒 FALSE。 *)
	aG2Valve : ARRAY[1..3] OF BOOL; (* G2 三个侧挡阀的电气电平 1=300，2=450，3=600；未接管时全 FALSE。 *)
	uiG2Band : UINT; (* G2 当前实际下降的料型带号 300/450/600；0 表示三缸全部提升，供诊断观察。 *)
END_VAR
VAR
	aConfig : ARRAY[1..17] OF ST_DeviceConfig; (* 设备配置数组，首扫描按固定编号设置类型和初始姿态。 *)
	aAxis : ARRAY[1..17] OF FB_Axis; (* 定位轴功能块实例数组，只有设备类型为 Axis 的元素被调用。 *)
	aMotor : ARRAY[1..17] OF FB_Motor; (* 连续电机功能块实例数组，供 D1、D3 使用。 *)
	aCylinder : ARRAY[1..17] OF FB_Cylinder; (* 气缸功能块实例数组，按 G 编号驱动对应仿真实例。 *)
	aValve : ARRAY[1..17] OF FB_Valve; (* 阀功能块实例数组，供 G5 喷油及 G6 吹气使用。 *)
	fbRealD1 : FB_RealAxis; (* D1 送料皮带真实轴实例，绑定 songliao。 *)
	fbRealD2 : FB_RealAxis; (* D2 切割走刀真实轴实例，绑定 qiege。 *)
	fbRealD3 : FB_RealAxis; (* D3 盘刀旋转真实轴实例，绑定 pandao（当前按线性模式配置）。 *)
	fbRealD8 : FB_RealAxis; (* D8 平台旋转真实轴实例，绑定 xuanzhuan（台达 ASDA-B3-E）。 *)
	fbRealG1 : FB_RealCylinder; (* G1 下压气缸真实实例，绑定左右两路阀与 G1 两端传感器。 *)
	fbRealG2 : FB_RealCylinderGroup; (* G2 侧挡气缸组真实实例，一台管 300/450/600 三个缸。 *)
	fbRealG3 : FB_RealCylinder; (* G3 侧推气缸真实实例，绑定 xDoG3Valve 与 G3 两端传感器。 *)
	fbRealG9 : FB_RealCylinder; (* G9 盘刀升降真实实例，绑定 xDoG9Valve 与 G9 两端传感器。 *)
	fbRealD6 : FB_RealSensor; (* D6 定长光电真实实例，只读；接管后取代 FB_SimPlant 产生料到位信号。 *)
	axUseReal : ARRAY[1..17] OF BOOL; (* 本扫描逐台接管标志，直接取 stReal.axRealDevice；没有真实实例的编号由回填分支报 3002。 *)
	xBooted : BOOL; (* 本功能块首次初始化完成标志，防止每扫描重写初值。 *)
	i : INT; (* 本扫描数组遍历索引；含义及范围以当前 FOR 循环为准。 *)
END_VAR

IF NOT xBooted THEN
	(* D1 送料皮带：由真实轴 songliao 承担输送，按定位轴建模（点动/连续运行）。 *)
	aConfig[1].eKind := E_DeviceKind.Axis;
	aConfig[2].eKind := E_DeviceKind.Axis;
	aConfig[3].eKind := E_DeviceKind.Motor;
	aConfig[4].eKind := E_DeviceKind.Axis;
	(* D5 暂按定位升降建模：0=升起避让，1=下降检测，非实际机械坐标。 *)
	aConfig[5].eKind := E_DeviceKind.Axis;
	aConfig[7].eKind := E_DeviceKind.Axis;
	aConfig[8].eKind := E_DeviceKind.Axis;
	FOR i := 9 TO 17 DO aConfig[i].eKind := E_DeviceKind.Cylinder; END_FOR
	aConfig[13].eKind := E_DeviceKind.Valve;
	aConfig[14].eKind := E_DeviceKind.Valve;
	aConfig[12].lrInitialPosition := 1.0;
	FOR i := 1 TO 17 DO
		IF aConfig[i].eKind = E_DeviceKind.Cylinder THEN
			aConfig[i].lrMinPosition := 0.0; aConfig[i].lrMaxPosition := 1.0;
		END_IF
	END_FOR
	(* D2 切割走刀：配方要求 200mm/s、加速度 500；默认 100/50 会把速度削到 100 并拖长加减速段。 *)
	aConfig[2].lrMaxVelocity := 300.0;
	aConfig[2].lrMaxAcceleration := 500.0;
	aConfig[2].lrMaxDeceleration := 500.0;
	xBooted := TRUE;
END_IF

(* 逐台接管标志直接取设置位：是否真的接管由下方回填分支的 CASE 决定。
   新增真实实例时只改 CASE 和实例调用两处，不要再维护第二份白名单。 *)
FOR i := 1 TO 17 DO
	axUseReal[i] := stReal.axRealDevice[i];
END_FOR

(* 四个真实轴实例每扫描必须无条件调用；轴形参写死，无法放进 FOR 循环。
   绑定对照（换电机、改轴名后必须逐行核对：写错不会报编译错误，
   因为任何一个合法轴名都能通过类型检查，只能靠单点测试发现）：
     fbRealD1 -> songliao    设备索引 1，送料皮带（EtherCAT 从站 ASDA_B3_E_CoE_Drive_3）
     fbRealD2 -> qiege       设备索引 2，切割走刀（从站 ASDA_B3_E_CoE_Drive_1）
     fbRealD3 -> pandao      设备索引 3，盘刀旋转（从站 ASDA_B3_E_CoE_Drive_2）
     fbRealD8 -> xuanzhuan   设备索引 8，平台旋转（从站 ASDA_B3_E_CoE_Drive，台达）
   注意：ASDA_B3_E_CoE_Drive_* 是驱动器从站名，代码里写的必须是它下面那个
   轴对象名（songliao/qiege/pandao/xuanzhuan），两者不是一回事。 *)
fbRealD1(Axis := songliao, xUseReal := axUseReal[1], xEnable := xEnable, xReset := xReset,
	xFaultHold := xFaultHold,
	stConfig := aConfig[1], stCommand := aCommand[1], stReal := stReal);
fbRealD2(Axis := qiege, xUseReal := axUseReal[2], xEnable := xEnable, xReset := xReset,
	xFaultHold := xFaultHold,
	stConfig := aConfig[2], stCommand := aCommand[2], stReal := stReal);
fbRealD3(Axis := pandao, xUseReal := axUseReal[3], xEnable := xEnable, xReset := xReset,
	xFaultHold := xFaultHold,
	stConfig := aConfig[3], stCommand := aCommand[3], stReal := stReal);
fbRealD8(Axis := xuanzhuan, xUseReal := axUseReal[8], xEnable := xEnable, xReset := xReset,
	xFaultHold := xFaultHold,
	stConfig := aConfig[8], stCommand := aCommand[8], stReal := stReal);

(* 四个真实气缸实例同样必须无条件调用；传感器与阀逐一对应物理映射符号。
   极性默认 FALSE：传感器高电平有效、阀高电平使能。接线反了只改这里一行，不动流程与互锁。 *)
fbRealG1(xUseReal := axUseReal[9], xEnable := xEnable, xReset := xReset,
	xFaultHold := xFaultHold,
	xSensorRetract := GVL_IO_Physical.xDiG1LRetract, xSensorExtend := GVL_IO_Physical.xDiG1LExtend,
	xSensorRetract2 := GVL_IO_Physical.xDiG1RRetract, xSensorExtend2 := GVL_IO_Physical.xDiG1RExtend,
	xUseSecond := TRUE,
	(* 现场 G1 两只伸出到位传感器已失效：改成只看左右两个缩回信号，两者都无信号并稳定 1s 即认为压到位。
	   传感器修好后把 xExtendByRetract 改回 FALSE 就恢复两端判定，流程和互锁都不用动。 *)
	xExtendByRetract := TRUE, tExtendConfirm := T#1S,
	xInvertSensors := FALSE, xInvertValve := FALSE,
	stConfig := aConfig[9], stCommand := aCommand[9]);
fbRealG2(xUseReal := axUseReal[10], xEnable := xEnable, xReset := xReset,
	xFaultHold := xFaultHold,
	uiMaterialModel := uiMaterialModel,
	xSensorRetract1 := GVL_IO_Physical.xDiG2_300Retract, xSensorExtend1 := GVL_IO_Physical.xDiG2_300Extend,
	xSensorRetract2 := GVL_IO_Physical.xDiG2_450Retract, xSensorExtend2 := GVL_IO_Physical.xDiG2_450Extend,
	xSensorRetract3 := GVL_IO_Physical.xDiG2_600Retract, xSensorExtend3 := GVL_IO_Physical.xDiG2_600Extend,
	xInvertSensors := FALSE, xInvertValve := FALSE,
	stConfig := aConfig[10], stCommand := aCommand[10]);
fbRealG3(xUseReal := axUseReal[11], xEnable := xEnable, xReset := xReset,
	xFaultHold := xFaultHold,
	xSensorRetract := GVL_IO_Physical.xDiG3Retract, xSensorExtend := GVL_IO_Physical.xDiG3Extend,
	xInvertSensors := FALSE, xInvertValve := FALSE,
	stConfig := aConfig[11], stCommand := aCommand[11]);
fbRealG9(xUseReal := axUseReal[17], xEnable := xEnable, xReset := xReset,
	xFaultHold := xFaultHold,
	xSensorRetract := GVL_IO_Physical.xDiG9Retract, xSensorExtend := GVL_IO_Physical.xDiG9Extend,
	xInvertSensors := FALSE, xInvertValve := FALSE,
	stConfig := aConfig[17], stCommand := aCommand[17]);

(* D6 定长光电：只读设备，没有阀也没有动作。
   接线极性反了改 xInvertSensor；光电抖动大改 tDebounce；不需要常亮/常灭监视就把 tStuckTimeout 置 T#0MS。 *)
fbRealD6(xUseReal := axUseReal[6], xEnable := xEnable, xReset := xReset,
	xSensorRaw := GVL_IO_Physical.xDiMaterialLength, xInvertSensor := FALSE,
	tDebounce := T#20MS, tStuckTimeout := T#0MS,
	stConfig := aConfig[6], stCommand := aCommand[6]);

(* 每周期按接管标志二选一：有真实实例的直接回填，否则按设备类型走仿真。
   「实例即事实」：本 CASE 列出全部已实现真实适配的编号，没列到的编号若置了接管位，
   就在 ELSE 分支明确报 3002，避免静默走仿真被误认为已接实机。 *)
(* G2 三个阀默认失电：只有走真实气缸组且缸确实在下降时才会被下面的 CASE 置位。 *)
aG2Valve[1] := FALSE; aG2Valve[2] := FALSE; aG2Valve[3] := FALSE;
uiG2Band := 0;
FOR i := 1 TO 17 DO
	aValveOut[i] := FALSE; aValveOutAux[i] := FALSE;
	IF axUseReal[i] THEN
		CASE i OF
		1: aStatus[i] := fbRealD1.stStatus;
		2: aStatus[i] := fbRealD2.stStatus;
		3: aStatus[i] := fbRealD3.stStatus;
		6: aStatus[i] := fbRealD6.stStatus;
		8: aStatus[i] := fbRealD8.stStatus;
		9: aStatus[i] := fbRealG1.stStatus; aValveOut[i] := fbRealG1.xValve; aValveOutAux[i] := fbRealG1.xValve2;
		10: aStatus[i] := fbRealG2.stStatus; aG2Valve := fbRealG2.aValve; uiG2Band := fbRealG2.uiActiveBand;
		11: aStatus[i] := fbRealG3.stStatus; aValveOut[i] := fbRealG3.xValve;
		17: aStatus[i] := fbRealG9.stStatus; aValveOut[i] := fbRealG9.xValve;
		ELSE
			(* 请求接管但本版本没有对应真实实例：只报错，不启动仿真，保持与老逻辑一致 *)
			aStatus[i].xError := TRUE;
			aStatus[i].udiErrorID := 3002;
		END_CASE
	ELSE
		CASE aConfig[i].eKind OF
		E_DeviceKind.Axis:
			aAxis[i](xSimulation:=xSimulation,xEnable:=xEnable,xReset:=xReset,
				xStall:=stSim.axStall[i],xInjectFault:=stSim.axFault[i],stConfig:=aConfig[i],stCommand:=aCommand[i]);
			aStatus[i] := aAxis[i].stStatus;
		E_DeviceKind.Motor:
			aMotor[i](xSimulation:=xSimulation,xEnable:=xEnable,xReset:=xReset,
				xStall:=stSim.axStall[i],xInjectFault:=stSim.axFault[i],stConfig:=aConfig[i],stCommand:=aCommand[i]);
			aStatus[i] := aMotor[i].stStatus;
		E_DeviceKind.Cylinder:
			aCylinder[i](xSimulation:=xSimulation,xEnable:=xEnable,xReset:=xReset,
				xStall:=stSim.axStall[i],xInjectFault:=stSim.axFault[i],stConfig:=aConfig[i],stCommand:=aCommand[i]);
			aStatus[i] := aCylinder[i].stStatus;
		E_DeviceKind.Valve:
			aValve[i](xSimulation:=xSimulation,xEnable:=xEnable,xReset:=xReset,
				xStall:=stSim.axStall[i],xInjectFault:=stSim.axFault[i],stConfig:=aConfig[i],stCommand:=aCommand[i]);
			aStatus[i] := aValve[i].stStatus;
		END_CASE
	END_IF
END_FOR

END_FUNCTION_BLOCK

// Device/Application/02_Devices/FB_Axis
(* 模块说明：定位轴适配入口。当前调用内部仿真；真实轴的 MC 功能块、回原点和限位尚未接入。 *)
FUNCTION_BLOCK FB_Axis
VAR_INPUT
    xSimulation : BOOL; (* TRUE 使用内部仿真；当前 FALSE 报未实现 3001，不会接管真实运动。 *)
    xEnable : BOOL; (* 本功能使能，电平有效；失能时不接受新的动作请求。 *)
    xReset : BOOL; (* 故障复位许可；仿真设备仅在故障注入已撤销时清除错误。 *)
    xStall : BOOL; (* 仿真卡住输入；TRUE 暂停位置推进且不发完成，保留忙状态。 *)
    xInjectFault : BOOL; (* 仿真设备故障输入；TRUE 锁存错误码 9001。 *)
    stConfig : ST_DeviceConfig; (* 设备类型、初始位置、软限位与仿真动作时间。 *)
    stCommand : ST_DeviceCommand; (* 当前单设备命令，含动作类型、序号、目标和速度。 *)
END_VAR
VAR_OUTPUT
    stStatus : ST_DeviceStatus; (* 本模块对外发布的状态；字段含义见其数据类型。 *)
END_VAR
VAR
    fbSimulation : FB_SimDevice; (* 内部设备仿真实例，真实设备适配尚未接入。 *)
END_VAR

(* 真实设备适配尚未接入；关闭仿真时返回 3001，避免误认为已具备实机控制。 *)
fbSimulation(xEnable := xEnable AND xSimulation, xReset := xReset,
    xStall := xStall, xInjectFault := xInjectFault,
    stConfig := stConfig, stCommand := stCommand);
stStatus := fbSimulation.stStatus;
IF NOT xSimulation THEN
    stStatus.xReady := FALSE; stStatus.xBusy := FALSE; stStatus.xActive := FALSE;
    stStatus.xError := TRUE; stStatus.udiErrorID := 3001;
END_IF

END_FUNCTION_BLOCK

// Device/Application/06_Simulation/FB_SimDevice
(* 模块说明：设备仿真模型：定位按固定时间插值、连续运行保持状态、点动按时间增量累计位置。 *)
FUNCTION_BLOCK FB_SimDevice
VAR_INPUT
    xEnable : BOOL; (* 本功能使能，电平有效；失能时不接受新的动作请求。 *)
    xReset : BOOL; (* 故障复位许可；仿真设备仅在故障注入已撤销时清除错误。 *)
    xStall : BOOL; (* 仿真卡住输入；TRUE 暂停位置推进且不发完成，保留忙状态。 *)
    xInjectFault : BOOL; (* 仿真设备故障输入；TRUE 锁存错误码 9001。 *)
    stConfig : ST_DeviceConfig; (* 设备类型、初始位置、软限位与仿真动作时间。 *)
    stCommand : ST_DeviceCommand; (* 当前单设备命令，含动作类型、序号、目标和速度。 *)
END_VAR
VAR_OUTPUT
    stStatus : ST_DeviceStatus; (* 本模块对外发布的状态；字段含义见其数据类型。 *)
END_VAR
VAR
    xBooted : BOOL; (* 本功能块首次初始化完成标志，防止每扫描重写初值。 *)
    xAction : BOOL; (* 仿真定时动作进行中；定位和建立连续运行状态使用，点动另行处理。 *)
    udiLastID : UDINT; (* 上次已接受序号，同一序号保持期间不重复启动动作。 *)
    lrStart : LREAL; (* 本次仿真定位的起始位置，用于按时间插值。 *)
    lrTarget : LREAL; (* 本次已接受定位命令的目标位置快照，用于时间插值。 *)
    lrJogDelta : LREAL; (* 点动相邻扫描的时间差，单位秒；速度乘该值取得本扫描位移。 *)
    tLastJog : TIME; (* 上扫描点动计时值，用于计算本扫描时间增量。 *)
    tonAction : TON; (* 仿真定位或建立连续运行状态的定时器。 *)
    tonJog : TON; (* 点动累计计时器，用于计算位置增量，设定计时上限 24 小时。 *)
END_VAR

(* 首次读取初始位置；以后位置由仿真动作累计，不在每周期重新归零。 *)
IF NOT xBooted THEN
    stStatus.lrPosition := stConfig.lrInitialPosition;
    xBooted := TRUE;
END_IF
IF xReset AND NOT xInjectFault THEN
    stStatus.xError := FALSE; stStatus.udiErrorID := 0;
END_IF
IF xInjectFault THEN 
	stStatus.xError := TRUE;
	stStatus.udiErrorID := 9001;
END_IF
stStatus.xReady := xEnable AND NOT stStatus.xError AND (stConfig.eKind <> E_DeviceKind.Unused);

(* 无许可、无请求或明确 Stop 时取消当前动作并清接收/完成序号。 *)
IF NOT stStatus.xReady OR (stCommand.eAction = E_DeviceAction.None)
   OR (stCommand.eAction = E_DeviceAction.Stop) THEN
    xAction := FALSE; udiLastID := 0;
    stStatus.xBusy := FALSE; stStatus.xActive := FALSE;
    stStatus.udiAcceptedID := 0; stStatus.udiCompletedID := 0;
(* 只接收不同于上次的非零序号；接收时检查速度与目标行程范围。 *)
ELSIF (stCommand.udiID <> 0) AND (stCommand.udiID <> udiLastID) THEN
    udiLastID := stCommand.udiID;
    stStatus.udiAcceptedID := udiLastID; stStatus.udiCompletedID := 0;
    lrStart := stStatus.lrPosition; lrTarget := stCommand.lrTarget;
    IF (ABS(stCommand.lrVelocity) > stConfig.lrMaxVelocity)
       OR ((stCommand.eAction = E_DeviceAction.Position) AND
           ((lrTarget < stConfig.lrMinPosition) OR (lrTarget > stConfig.lrMaxPosition))) THEN
        stStatus.xError := TRUE; stStatus.udiErrorID := 2001; xAction := FALSE;
    ELSE
        xAction := stCommand.eAction <> E_DeviceAction.Jog;
        stStatus.xBusy := TRUE; stStatus.xActive := FALSE;
    END_IF
    (* 接收新序号时先复位计时器，随后由每扫描调用开始本次计时。 *)
    tonAction(IN := FALSE);
END_IF
(* 固定时间仿真定位，不依据实际速度/加速度建模；卡住注入时保持忙且不完成。 *)
tonAction(IN := xAction AND stStatus.xReady, PT := stConfig.tSimAction);
IF xAction AND NOT xStall AND stStatus.xReady THEN
    IF stCommand.eAction = E_DeviceAction.Position THEN
        stStatus.lrPosition := lrStart + (lrTarget-lrStart) *
            MIN(1.0, TIME_TO_LREAL(tonAction.ET) / MAX(1.0, TIME_TO_LREAL(stConfig.tSimAction)));
    END_IF
    IF tonAction.Q THEN
        IF stCommand.eAction = E_DeviceAction.Position THEN stStatus.lrPosition := lrTarget; END_IF
        stStatus.xBusy := FALSE;
        stStatus.xActive := stCommand.eAction = E_DeviceAction.Run;
        stStatus.udiCompletedID := udiLastID;
        xAction := FALSE;
    END_IF
END_IF
(* 点动按相邻扫描的时间差累计位置，达到示例软行程边界后限幅。 *)
tonJog(IN := stStatus.xReady AND (stCommand.eAction = E_DeviceAction.Jog), PT := T#24H);
IF tonJog.IN THEN
    lrJogDelta := TIME_TO_LREAL(tonJog.ET-tLastJog) / 1000.0;
    IF NOT xStall THEN
        stStatus.lrPosition := LIMIT(stConfig.lrMinPosition,
            stStatus.lrPosition+stCommand.lrVelocity*lrJogDelta, stConfig.lrMaxPosition);
    END_IF
    stStatus.xBusy := TRUE; stStatus.xActive := TRUE;
    tLastJog := tonJog.ET;
ELSE tLastJog := T#0MS;
END_IF
IF stStatus.xError THEN
    stStatus.xReady := FALSE; stStatus.xBusy := FALSE; stStatus.xActive := FALSE;
END_IF

END_FUNCTION_BLOCK

// Device/Application/02_Devices/FB_Motor
(* 模块说明：连续电机适配入口，供皮带 D1 和盘刀 D3 使用。当前仅仿真运行状态。 *)
FUNCTION_BLOCK FB_Motor
VAR_INPUT
    xSimulation : BOOL; (* TRUE 使用内部仿真；当前 FALSE 报未实现 3001，不会接管真实运动。 *)
    xEnable : BOOL; (* 本功能使能，电平有效；失能时不接受新的动作请求。 *)
    xReset : BOOL; (* 故障复位许可；仿真设备仅在故障注入已撤销时清除错误。 *)
    xStall : BOOL; (* 仿真卡住输入；TRUE 暂停位置推进且不发完成，保留忙状态。 *)
    xInjectFault : BOOL; (* 仿真设备故障输入；TRUE 锁存错误码 9001。 *)
    stConfig : ST_DeviceConfig; (* 设备类型、初始位置、软限位与仿真动作时间。 *)
    stCommand : ST_DeviceCommand; (* 当前单设备命令，含动作类型、序号、目标和速度。 *)
END_VAR
VAR_OUTPUT
    stStatus : ST_DeviceStatus; (* 本模块对外发布的状态；字段含义见其数据类型。 *)
END_VAR
VAR
    fbSimulation : FB_SimDevice; (* 内部设备仿真实例，真实设备适配尚未接入。 *)
END_VAR

(* 真实设备适配尚未接入；关闭仿真时返回 3001，避免误认为已具备实机控制。 *)
fbSimulation(xEnable := xEnable AND xSimulation, xReset := xReset,
    xStall := xStall, xInjectFault := xInjectFault,
    stConfig := stConfig, stCommand := stCommand);
stStatus := fbSimulation.stStatus;
IF NOT xSimulation THEN
    stStatus.xReady := FALSE; stStatus.xBusy := FALSE; stStatus.xActive := FALSE;
    stStatus.xError := TRUE; stStatus.udiErrorID := 3001;
END_IF

END_FUNCTION_BLOCK

// Device/Application/02_Devices/FB_Cylinder
(* 模块说明：气缸适配入口。当前用 0/1 位置模拟两端到位；真实电磁阀和到位传感器尚未映射。 *)
FUNCTION_BLOCK FB_Cylinder
VAR_INPUT
    xSimulation : BOOL; (* TRUE 使用内部仿真；当前 FALSE 报未实现 3001，不会接管真实运动。 *)
    xEnable : BOOL; (* 本功能使能，电平有效；失能时不接受新的动作请求。 *)
    xReset : BOOL; (* 故障复位许可；仿真设备仅在故障注入已撤销时清除错误。 *)
    xStall : BOOL; (* 仿真卡住输入；TRUE 暂停位置推进且不发完成，保留忙状态。 *)
    xInjectFault : BOOL; (* 仿真设备故障输入；TRUE 锁存错误码 9001。 *)
    stConfig : ST_DeviceConfig; (* 设备类型、初始位置、软限位与仿真动作时间。 *)
    stCommand : ST_DeviceCommand; (* 当前单设备命令，含动作类型、序号、目标和速度。 *)
END_VAR
VAR_OUTPUT
    stStatus : ST_DeviceStatus; (* 本模块对外发布的状态；字段含义见其数据类型。 *)
END_VAR
VAR
    fbSimulation : FB_SimDevice; (* 内部设备仿真实例，真实设备适配尚未接入。 *)
END_VAR

(* 真实设备适配尚未接入；关闭仿真时返回 3001，避免误认为已具备实机控制。 *)
fbSimulation(xEnable := xEnable AND xSimulation, xReset := xReset,
    xStall := xStall, xInjectFault := xInjectFault,
    stConfig := stConfig, stCommand := stCommand);
stStatus := fbSimulation.stStatus;
IF NOT xSimulation THEN
    stStatus.xReady := FALSE; stStatus.xBusy := FALSE; stStatus.xActive := FALSE;
    stStatus.xError := TRUE; stStatus.udiErrorID := 3001;
END_IF

END_FUNCTION_BLOCK

// Device/Application/02_Devices/FB_Valve
(* 模块说明：阀适配入口，供喷油 G5 和吹气 G6 使用。当前用运行状态表示开启，未映射输出。 *)
FUNCTION_BLOCK FB_Valve
VAR_INPUT
    xSimulation : BOOL; (* TRUE 使用内部仿真；当前 FALSE 报未实现 3001，不会接管真实运动。 *)
    xEnable : BOOL; (* 本功能使能，电平有效；失能时不接受新的动作请求。 *)
    xReset : BOOL; (* 故障复位许可；仿真设备仅在故障注入已撤销时清除错误。 *)
    xStall : BOOL; (* 仿真卡住输入；TRUE 暂停位置推进且不发完成，保留忙状态。 *)
    xInjectFault : BOOL; (* 仿真设备故障输入；TRUE 锁存错误码 9001。 *)
    stConfig : ST_DeviceConfig; (* 设备类型、初始位置、软限位与仿真动作时间。 *)
    stCommand : ST_DeviceCommand; (* 当前单设备命令，含动作类型、序号、目标和速度。 *)
END_VAR
VAR_OUTPUT
    stStatus : ST_DeviceStatus; (* 本模块对外发布的状态；字段含义见其数据类型。 *)
END_VAR
VAR
    fbSimulation : FB_SimDevice; (* 内部设备仿真实例，真实设备适配尚未接入。 *)
END_VAR

(* 真实设备适配尚未接入；关闭仿真时返回 3001，避免误认为已具备实机控制。 *)
fbSimulation(xEnable := xEnable AND xSimulation, xReset := xReset,
    xStall := xStall, xInjectFault := xInjectFault,
    stConfig := stConfig, stCommand := stCommand);
stStatus := fbSimulation.stStatus;
IF NOT xSimulation THEN
    stStatus.xReady := FALSE; stStatus.xBusy := FALSE; stStatus.xActive := FALSE;
    stStatus.xError := TRUE; stStatus.udiErrorID := 3001;
END_IF

END_FUNCTION_BLOCK

// Device/Application/02_Devices/FB_RealAxis
FUNCTION_BLOCK FB_RealAxis
(* 模块说明：真实轴适配层。把统一设备命令翻译成 SoftMotion 动作，并回写与仿真完全一致的接收/完成序号。 *)
VAR_IN_OUT
	Axis : AXIS_REF_SM3; (* 轴节点引用，编译期强制绑定；未接轴无法通过编译，不存在空指针。 *)
END_VAR
VAR_INPUT
	xUseReal : BOOL; (* TRUE 表示本编号由本功能块接管；FALSE 时驱动器保持去使能且不响应任何命令。 *)
	xEnable : BOOL; (* 设备级使能，来自整机许可；FALSE 时主动停止并清序号。 *)
	xReset : BOOL; (* 故障复位，上升沿清锁存错误与 MC 错误。 *)
	stConfig : ST_DeviceConfig; (* 行程、速度、加减速与绝对定位许可。 *)
	stCommand : ST_DeviceCommand; (* 上层统一设备命令，含义与仿真侧完全一致。 *)
	xFaultHold : BOOL; (* 整机故障保持：TRUE 期间强制 MC_Stop 常置并清所有运动请求，直到复位。 *)
	stReal : ST_RealDeviceSettings; (* 相对验证距离、速度与旁路设置。 *)
END_VAR
VAR_OUTPUT
	stStatus : ST_DeviceStatus; (* 与 FB_SimDevice 语义一致，上层无需区分真假设备。 *)
	uiVerifyPhase : UINT; (* 相对验证相位：0 空闲、1 正向、2 停留、3 反向、4 完成、90 中止。 *)
	lrVerifyMeasured : LREAL; (* 本次往返正向段的实测位移，取自轴反馈。 *)
	lrVerifyRatio : LREAL; (* 实测除以指令；只能证明指令与反馈自洽，不能证明单位就是毫米。 *)
END_VAR
VAR
	fbPower : MC_Power; (* 伺服使能，接管期间保持上电。 *)
	fbReset : MC_Reset; (* 清 MC 错误。 *)
	fbStop : MC_Stop; (* 受控停止，停止请求需保持到 Done。 *)
	fbMoveAbs : MC_MoveAbsolute; (* 绝对定位，仅在 xAbsoluteAllowed 为 TRUE 时使用。 *)
	fbMoveRel : MC_MoveRelative; (* 相对定位，验证模式的两段行程使用。 *)
	fbMoveVel : MC_MoveVelocity; (* 连续运行与点动共用，两者相位互斥；方向必须显式给出。 *)
	fbHoming : CmpHCMotion.MC_Homing; (* 上位机回零：由 PLC 自己按轴配置的回零方式走，不依赖驱动器支持 DS402 回零。 *)
	fbReadPos : MC_ReadActualPosition; (* 实际位置反馈。 *)
	fbReadStatus : MC_ReadStatus; (* 轴状态，用于判断故障停止。 *)
	fbReadErr : MC_ReadAxisError; (* 轴错误码，供在线排查。 *)
	rtReset : R_TRIG; (* 复位上升沿。 *)
	tonEnable : TON; (* 命令已接收但轴未使能的 3 秒超时。 *)
	tonDwell : TON; (* 验证往返之间的停留，保证 Execute 拉低形成新上升沿。 *)
	tonHome : TON; (* 回零超时；找不到原点时按 2004 暴露，避免无限等待。 *)
	udiLastID : UDINT; (* 上次已接受序号，用于识别新命令。 *)
	udiActiveID : UDINT; (* 正在执行的序号，完成时回写。 *)
	xPending : BOOL; (* 已接收但尚未启动，等待轴使能。 *)
	xStopLatch : BOOL; (* 停止请求锁存，保持到 MC_Stop 完成。 *)
	xStopReq : BOOL; (* 本扫描停止请求。 *)
	xMoveAbsReq : BOOL; (* 本扫描绝对定位请求。 *)
	xMoveRelReq : BOOL; (* 本扫描相对定位请求。 *)
	xMoveVelReq : BOOL; (* 本扫描速度模式请求，连续运行与点动共用。 *)
	xHomeReq : BOOL; (* 本扫描回零请求，保持到 Done。 *)
	xHomed : BOOL; (* 本次上电后已成功回零；成功后允许绝对定位，断电或重新下载后清零。 *)
	uiPhase : UINT; (* 动作相位：0 空闲、10 等待使能、20 绝对、30/31/32 验证三段、40 连续、50 点动、60 回零、90 中止。 *)
	lrVerifyStart : LREAL; (* 验证正向段起点位置。 *)
	lrRelDistance : LREAL; (* 本次相对定位距离，正负决定方向。 *)
	lrRelVelocity : LREAL; (* 本次相对定位速度，取正值。 *)
	lrCmdVelocity : LREAL; (* 连续运行与点动的限幅后速度，带符号。 *)
END_VAR

(* ===== 1. 读取块无条件调用，保证反馈新鲜 ===== *)
fbReadPos(Axis := Axis, Enable := TRUE);
fbReadStatus(Axis := Axis, Enable := TRUE);
fbReadErr(Axis := Axis, Enable := TRUE);
rtReset(CLK := xReset);

stStatus.lrPosition := fbReadPos.Position;
stStatus.xRealActive := xUseReal;

(* ===== 2. 复位：只在接管状态下响应，避免误清其它轴 ===== *)
IF xUseReal AND rtReset.Q THEN
	stStatus.xError := FALSE;
	stStatus.udiErrorID := 0;
	xStopLatch := FALSE;
	xPending := FALSE;
	uiPhase := 0;
	uiVerifyPhase := 0;
	udiLastID := 0;
	udiActiveID := 0;
	stStatus.udiAcceptedID := 0;
	stStatus.udiCompletedID := 0;
	stStatus.xBusy := FALSE;
	stStatus.xActive := FALSE;
END_IF

(* ===== 3. 定时器：用上扫描状态驱动，避免与状态判定循环依赖 ===== *)
tonEnable(IN := xPending AND xUseReal, PT := T#3S);
tonDwell(IN := (uiPhase = 31), PT := stReal.tVerifyDwell);
tonHome(IN := (uiPhase = 60), PT := stReal.tHomeTimeout);

(* ===== 4. 请求默认全部撤销 ===== *)
xStopReq := FALSE;
xMoveAbsReq := FALSE;
xMoveRelReq := FALSE;
xMoveVelReq := FALSE;
xHomeReq := FALSE;
lrRelDistance := 0.0;
lrRelVelocity := 0.0;
lrCmdVelocity := 0.0;

(* ===== 4.5 整机故障保持：故障期间主动停车，不依赖 xPermit 间接撤销 ===== *)
(* 为什么需要：进入 Fault 时上层只是让 xPermit 变 FALSE，请求被换成 Stop。但 Stop 是
   一次性的动作请求，盘刀这类连续运行设备在 MC_Stop 完成后再无后续指令，表现就是
   “PLC 认为已停、实际还在转”。这里改用 xFaultHold 强制 MC_Stop 常置，直到真正复位。 *)
IF xFaultHold THEN
	xStopReq := TRUE;
	xPending := FALSE;
	xMoveAbsReq := FALSE; xMoveRelReq := FALSE; xMoveVelReq := FALSE; xHomeReq := FALSE;
	uiPhase := 0; uiVerifyPhase := 0;
	udiLastID := 0; udiActiveID := 0;
	stStatus.udiAcceptedID := 0; stStatus.udiCompletedID := 0;
	stStatus.xBusy := FALSE; stStatus.xActive := FALSE;
END_IF

(* ===== 5. 主状态判定 ===== *)
IF NOT xUseReal THEN
	(* 未接管：不产生任何运动请求，驱动器由 MC_Power 去使能。 *)
	xPending := FALSE; xStopLatch := FALSE;
	uiPhase := 0; uiVerifyPhase := 0;
	udiLastID := 0; udiActiveID := 0;
	stStatus.xReady := FALSE;
	stStatus.xBusy := FALSE; stStatus.xActive := FALSE;
	stStatus.udiAcceptedID := 0; stStatus.udiCompletedID := 0;
	stStatus.xError := FALSE; stStatus.udiErrorID := 0;
ELSIF xFaultHold THEN
	(* 故障保持：只允许停止，不接收新命令，也不发布就绪。 *)
	stStatus.xReady := FALSE;
	stStatus.xBusy := FALSE; stStatus.xActive := FALSE;
	stStatus.udiAcceptedID := 0; stStatus.udiCompletedID := 0;
ELSE
	(* --- 5.1 接收新序号：新序号就是新命令，不用边沿检测 --- *)
	IF (stCommand.udiID <> 0) AND (stCommand.udiID <> udiLastID)
		AND xEnable AND NOT stStatus.xError THEN
		udiLastID := stCommand.udiID;
		udiActiveID := udiLastID;
		stStatus.udiAcceptedID := udiActiveID;
		stStatus.udiCompletedID := 0;
		stStatus.xBusy := TRUE; stStatus.xActive := FALSE;
		uiVerifyPhase := 0;
		xPending := TRUE;
		uiPhase := 10;
		xStopLatch := FALSE;
	END_IF

	(* --- 5.2 停止请求锁存：保持到 MC_Stop 完成，不能提前撤 Execute --- *)
	IF (stCommand.eAction = E_DeviceAction.Stop) OR (NOT xEnable) THEN
		(* 只在真的有动作时才锁存，避免 Stop 常驻时每扫描重复触发 MC_Stop。 *)
		IF xPending OR (uiPhase <> 0) THEN xStopLatch := TRUE; END_IF
	ELSIF (stCommand.eAction = E_DeviceAction.None) AND (uiPhase <> 0) THEN
		xStopLatch := TRUE;
	END_IF
	IF fbStop.Done THEN xStopLatch := FALSE; END_IF

	IF xStopLatch THEN
		xStopReq := TRUE;
		xPending := FALSE;
		uiPhase := 0; uiVerifyPhase := 0;
		udiLastID := 0; udiActiveID := 0;
		stStatus.udiAcceptedID := 0; stStatus.udiCompletedID := 0;
		stStatus.xBusy := FALSE; stStatus.xActive := FALSE;
	ELSIF xPending THEN
		(* --- 5.3 等轴使能；就绪后按动作类型进入相位，3 秒未使能报 2003 --- *)
		IF fbPower.Status THEN
			xPending := FALSE;
			CASE stCommand.eAction OF
			E_DeviceAction.Position:
				(* 已回零优先走绝对定位：相对验证只是未回零时的临时替代，回零成功后不再需要。 *)
				IF xHomed OR stConfig.xAbsoluteAllowed THEN
					uiPhase := 20;
				ELSIF stReal.xRelativeVerify THEN
					lrVerifyStart := fbReadPos.Position;
					uiPhase := 30; uiVerifyPhase := 1;
				ELSE
					(* 未回零不允许绝对定位：报 2002 且不置完成位，由上层按步号超时暴露。 *)
					stStatus.xError := TRUE; stStatus.udiErrorID := 2002;
					uiPhase := 0; uiVerifyPhase := 0;
				END_IF
			E_DeviceAction.Run:
				uiPhase := 40;
			E_DeviceAction.Jog:
				uiPhase := 50;
			E_DeviceAction.Home:
				uiPhase := 60;
			ELSE
				uiPhase := 0;
			END_CASE
		ELSIF tonEnable.Q THEN
			xPending := FALSE; uiPhase := 0;
			stStatus.xError := TRUE; stStatus.udiErrorID := 2003;
			stStatus.xBusy := FALSE;
		END_IF
	END_IF

	(* --- 5.4 按相位生成限幅后的运动参数 --- *)
	CASE uiPhase OF
	30:
		lrRelDistance := LIMIT(0.0, stReal.lrVerifyDistance, 20.0);
		lrRelVelocity := LIMIT(0.01, stReal.lrVerifyVelocity, stConfig.lrMaxVelocity);
	32:
		lrRelDistance := -LIMIT(0.0, stReal.lrVerifyDistance, 20.0);
		lrRelVelocity := LIMIT(0.01, stReal.lrVerifyVelocity, stConfig.lrMaxVelocity);
	40:
		(* 连续运行：按设备配置限幅，不使用验证低速。 *)
		lrCmdVelocity := LIMIT(-stConfig.lrMaxVelocity, stCommand.lrVelocity, stConfig.lrMaxVelocity);
	50:
		(* 点动：用设备最大速度与手动上限 lrManualVelocityMax 的较小者限幅；不能再用验证速度，否则手动最高只有 2mm/s。 *)
		lrCmdVelocity := LIMIT(0.01, ABS(stCommand.lrVelocity),
			MIN(stConfig.lrMaxVelocity, stReal.lrManualVelocityMax));
		IF stCommand.lrVelocity < 0.0 THEN lrCmdVelocity := -lrCmdVelocity; END_IF
	END_CASE

	xMoveAbsReq := (uiPhase = 20);
	xMoveRelReq := (uiPhase = 30) OR (uiPhase = 32);
	xMoveVelReq := (uiPhase = 40) OR (uiPhase = 50);
	xHomeReq := (uiPhase = 60);
END_IF

(* ===== 6. MC 块无条件调用：漏调用会报 SMC_FB_WASNT_CALLED_DURING_MOTION ===== *)
fbPower(Axis := Axis, Enable := xUseReal AND xEnable,
	bRegulatorOn := xUseReal AND xEnable, bDriveStart := xUseReal AND xEnable);
fbReset(Axis := Axis, Execute := xUseReal AND rtReset.Q);
fbStop(Axis := Axis, Execute := xStopReq OR xFaultHold, Deceleration := stConfig.lrMaxDeceleration);
fbMoveRel(Axis := Axis, Execute := xMoveRelReq, Distance := lrRelDistance,
	Velocity := lrRelVelocity, Acceleration := stConfig.lrMaxAcceleration,
	Deceleration := stConfig.lrMaxDeceleration);
fbMoveAbs(Axis := Axis, Execute := xMoveAbsReq, Position := stCommand.lrTarget,
	Velocity := LIMIT(0.01, ABS(stCommand.lrVelocity), stConfig.lrMaxVelocity),
	Acceleration := stConfig.lrMaxAcceleration, Deceleration := stConfig.lrMaxDeceleration);
fbMoveVel(Axis := Axis, Execute := xMoveVelReq,
	Velocity := ABS(lrCmdVelocity),
	Direction := SEL(lrCmdVelocity < 0.0, MC_Direction.positive, MC_Direction.negative),
	Acceleration := stConfig.lrMaxAcceleration,
	Deceleration := stConfig.lrMaxDeceleration);
(* 回零走 MC_Homing（上位机回零）：回零方式、开始方向、零点信号、快慢速全部来自轴配置，
   本块只给 Axis 和 Execute。驱动器不支持 DS402 回零，用 MC_Home 会一直卡在 Homing 状态不动。 *)
fbHoming(Axis := Axis, Execute := xHomeReq);

(* ===== 7. 完成判定与序号回写 ===== *)
IF xUseReal THEN
	CASE uiPhase OF
	20:
		IF fbMoveAbs.Done THEN
			stStatus.udiCompletedID := udiActiveID;
			stStatus.xBusy := FALSE; stStatus.xActive := FALSE;
			uiPhase := 0;
		ELSIF fbMoveAbs.CommandAborted THEN
			stStatus.xBusy := FALSE; uiPhase := 0;
		END_IF
	30:
		IF fbMoveRel.Done THEN
			lrVerifyMeasured := fbReadPos.Position - lrVerifyStart;
			uiPhase := 31; uiVerifyPhase := 2;
		ELSIF fbMoveRel.CommandAborted THEN
			uiPhase := 90; uiVerifyPhase := 90;
			stStatus.xError := TRUE; stStatus.udiErrorID := 2005;
			stStatus.xBusy := FALSE;
		END_IF
	31:
		IF tonDwell.Q THEN
			uiPhase := 32; uiVerifyPhase := 3;
		END_IF
	32:
		IF fbMoveRel.Done THEN
			IF stReal.lrVerifyDistance > 0.001 THEN
				lrVerifyRatio := lrVerifyMeasured / stReal.lrVerifyDistance;
			END_IF
			uiPhase := 0; uiVerifyPhase := 4;
			stStatus.udiCompletedID := udiActiveID;
			stStatus.xBusy := FALSE; stStatus.xActive := FALSE;
		ELSIF fbMoveRel.CommandAborted THEN
			uiPhase := 90; uiVerifyPhase := 90;
			stStatus.xError := TRUE; stStatus.udiErrorID := 2005;
			stStatus.xBusy := FALSE;
		END_IF
	40:
		(* 连续运行：建立速度后回写完成位，但保持相位直到命令改变。 *)
		IF fbMoveVel.InVelocity THEN
			stStatus.xActive := TRUE;
			stStatus.xBusy := FALSE;
			stStatus.udiCompletedID := udiActiveID;
		END_IF
	50:
		(* 点动：与仿真一致，不置完成位，靠松开后的 None/Stop 停止。 *)
		stStatus.xActive := fbMoveVel.InVelocity;
		stStatus.xBusy := TRUE;
	60:
		(* 回零：Done 后置 xHomed 并放行绝对定位；超时报 2004 且不置完成位，避免上层误判已到位。 *)
		IF fbHoming.Done THEN
			xHomed := TRUE;
			stStatus.udiCompletedID := udiActiveID;
			stStatus.xBusy := FALSE; stStatus.xActive := FALSE;
			uiPhase := 0;
		ELSIF fbHoming.CommandAborted THEN
			(* 被其它运动块打断：只清忙标志退出相位，既不置完成位也不置故障，由上层按步号超时暴露。 *)
			stStatus.xBusy := FALSE; uiPhase := 0;
		ELSIF tonHome.Q THEN
			xHomed := FALSE;
			stStatus.xError := TRUE; stStatus.udiErrorID := 2004;
			stStatus.xBusy := FALSE; uiPhase := 0;
		END_IF
	END_CASE

	(* --- MC 错误汇总：只锁存第一条，40000 为前缀，低 16 位保留原码便于查手册 --- *)
	IF NOT stStatus.xError THEN
		IF fbPower.Error THEN
			stStatus.xError := TRUE; stStatus.udiErrorID := UDINT#40000 + TO_UDINT(fbPower.ErrorID);
		ELSIF fbReset.Error THEN
			stStatus.xError := TRUE; stStatus.udiErrorID := UDINT#40000 + TO_UDINT(fbReset.ErrorID);
		ELSIF fbStop.Error THEN
			stStatus.xError := TRUE; stStatus.udiErrorID := UDINT#40000 + TO_UDINT(fbStop.ErrorID);
		ELSIF fbMoveRel.Error THEN
			stStatus.xError := TRUE; stStatus.udiErrorID := UDINT#40000 + TO_UDINT(fbMoveRel.ErrorID);
		ELSIF fbMoveAbs.Error THEN
			stStatus.xError := TRUE; stStatus.udiErrorID := UDINT#40000 + TO_UDINT(fbMoveAbs.ErrorID);
		ELSIF fbMoveVel.Error THEN
			stStatus.xError := TRUE; stStatus.udiErrorID := UDINT#40000 + TO_UDINT(fbMoveVel.ErrorID);
		ELSIF fbHoming.Error THEN
			stStatus.xError := TRUE; stStatus.udiErrorID := UDINT#40000 + TO_UDINT(fbHoming.ErrorID);
		END_IF
	END_IF
END_IF

(* ===== 8. 就绪与故障收尾 ===== *)
stStatus.xReady := xUseReal AND xEnable AND NOT stStatus.xError;
stStatus.xHomed := xUseReal AND xHomed;
IF stStatus.xError THEN
	stStatus.xBusy := FALSE;
	stStatus.xActive := FALSE;
END_IF

END_FUNCTION_BLOCK

// Device/Application/02_Devices/FB_RealCylinder
FUNCTION_BLOCK FB_RealCylinder
(* 模块说明：真实气缸适配层。读取两端到位传感器判定姿态，按统一设备命令驱动单电控阀，
   回写与 FB_SimDevice 完全一致的接收/完成序号，使上层流程与互锁无需区分真假气缸。
   某个端点传感器损坏时用 xExtendByRetract 退让：只看缩回信号，全部消失并稳定后视为伸出到位。 *)
VAR_INPUT
	xUseReal : BOOL; (* TRUE 表示本编号由真实气缸接管；FALSE 时阀保持失电且不响应任何命令。 *)
	xEnable : BOOL; (* 设备级使能，来自整机许可；FALSE 时阀失电并清序号。 *)
	xReset : BOOL; (* 故障复位上升沿；清锁存错误并允许重新建立姿态。 *)
	xSensorRetract : BOOL; (* 缩回到位传感器原始电平，TRUE 表示该端有信号。 *)
	xSensorExtend : BOOL; (* 伸出到位传感器原始电平，TRUE 表示该端有信号。 *)
	xSensorRetract2 : BOOL; (* 第二组（右压板）缩回到位原始电平；仅 xUseSecond 为 TRUE 时参与判定。 *)
	xSensorExtend2 : BOOL; (* 第二组（右压板）伸出到位原始电平；仅 xUseSecond 为 TRUE 时参与判定。 *)
	xUseSecond : BOOL := FALSE; (* TRUE 表示由两个同步执行器组成：两组传感器必须同时到位才算该端到位。 *)
	xExtendByRetract : BOOL := FALSE; (* 退让模式：伸出端传感器不可用时置 TRUE，改用「所有缩回信号都消失」推断伸出到位；默认 FALSE 仍按两端判定。 *)
	tExtendConfirm : TIME := T#1S; (* 仅退让模式有效：缩回信号消失并持续该时间才确认伸出到位，避免气缸刚起步就误判为已伸出。 *)
	xInvertSensors : BOOL; (* TRUE 表示两个传感器接线为低电平有效，本层统一取反，不动上层。 *)
	xInvertValve : BOOL; (* TRUE 表示阀为低电平使能；默认 FALSE，即高电平使能。 *)
	xFaultHold : BOOL := FALSE; (* 整机故障保持：TRUE 时阀立即失电并撤销保位，直到复位。 *)
	tSensorTimeout : TIME := T#3S; (* 两端均无信号达到该时间判为传感器丢失，报 3004；双执行器时也包含两侧不同步。 *)
	tTravelTimeout : TIME := T#10S; (* 命令发出后未到位达到该时间判为动作超时，报 3005。 *)
	stConfig : ST_DeviceConfig; (* 行程范围，语义与仿真侧一致；气缸只使用 0/1 两端。 *)
	stCommand : ST_DeviceCommand; (* 上层统一设备命令，气缸只响应 Position 的 0/1 目标。 *)
END_VAR
VAR_OUTPUT
	stStatus : ST_DeviceStatus; (* 与 FB_SimDevice 语义一致；lrPosition 取 0.0 缩回、1.0 伸出。 *)
	xValve : BOOL; (* 阀电气输出电平，已含 xInvertValve；直接接物理输出点。 *)
	xValve2 : BOOL; (* 第二个执行器的阀电气输出电平；xUseSecond 为 FALSE 时恒为 FALSE。 *)
END_VAR
VAR
	rtReset : R_TRIG; (* 复位上升沿。 *)
	tonNoSensor : TON; (* 两端均无信号的持续计时。 *)
	tonExtendConfirm : TON; (* 退让模式下「缩回信号全部消失」的持续计时，到时才确认伸出到位。 *)
	tonTravel : TON; (* 命令发出后等待到位的计时。 *)
	udiLastID : UDINT; (* 上次已接受的命令序号。 *)
	xSenseRetract : BOOL; (* 取反处理后的缩回信号：双执行器时为两侧 AND，TRUE 表示两侧都缩回到位。 *)
	xRetractAny : BOOL; (* 取反处理后的缩回信号：双执行器时为两侧 OR，TRUE 表示至少一侧仍停在缩回位。退让模式用它判「两侧都离开」。 *)
	xSenseExtend : BOOL; (* 取反处理后的伸出信号。 *)
	xPositionKnown : BOOL; (* 姿态是否已由传感器确立；未确立时 xReady 必须为 FALSE，防止上层把未知当成已缩回。 *)
	lrLastKnown : LREAL; (* 最后一次确立的姿态；传感器全灭时保持该值。 *)
	xCmdValid : BOOL; (* 当前存在有效的保位命令，阀按此持续输出。 *)
	xCmdExtend : BOOL; (* 有效命令期望的端点：TRUE 伸出，FALSE 缩回。 *)
	xTravelling : BOOL; (* 尚未确认到达目标端点。 *)
END_VAR

rtReset(CLK := xReset);

(* ===== 1. 复位：只清错误与序号，姿态仍由传感器决定 ===== *)
IF xUseReal AND rtReset.Q THEN
	stStatus.xError := FALSE; stStatus.udiErrorID := 0;
	xCmdValid := FALSE; xTravelling := FALSE; udiLastID := 0;
	stStatus.udiAcceptedID := 0; stStatus.udiCompletedID := 0;
	tonNoSensor(IN := FALSE);
	tonTravel(IN := FALSE);
END_IF

(* ===== 2. 传感器取反与姿态判定 ===== *)
xSenseRetract := xSensorRetract XOR xInvertSensors;
xSenseExtend := xSensorExtend XOR xInvertSensors;

(* 双执行器：两组必须同时到位才算该端到位。
   左侧在上、右侧在下时两个都为 FALSE，自然落进下面的“两端都无信号”分支：
   保持上次姿态，持续 tSensorTimeout 才报 3004，与单缸中间态同一套处理。
   同时另算一个 OR 合成量给退让模式用：AND 取反只能得到「至少一侧离开」，
   而退让模式要的是「两侧都离开」，所以必须在合并之前留一份单侧信号。 *)
xRetractAny := xSenseRetract;
IF xUseSecond THEN
	xRetractAny := xRetractAny OR (xSensorRetract2 XOR xInvertSensors);
	xSenseRetract := xSenseRetract AND (xSensorRetract2 XOR xInvertSensors);
	xSenseExtend := xSenseExtend AND (xSensorExtend2 XOR xInvertSensors);
END_IF

(* 退让模式：伸出端传感器不可用，只认缩回信号。
   判定 = 左右两侧都没有缩回信号（都离开缩回位）并持续 tExtendConfirm；
   必须延时确认：缩回信号在气缸刚起步就掉，不延时会在压板还没压下去时就报已伸出，
   上层的压紧判定和自动流程会提前放行。延时期间保持上次姿态。 *)
tonExtendConfirm(IN := xUseReal AND xExtendByRetract AND NOT xRetractAny, PT := tExtendConfirm);
IF xExtendByRetract THEN
	xSenseExtend := tonExtendConfirm.Q;
END_IF

(* 退让模式下「两端都无信号」正是伸出到位的正常表现，不能再按传感器丢失报 3004，所以此模式关闭该计时。 *)
tonNoSensor(IN := xUseReal AND NOT xExtendByRetract AND NOT xSenseRetract AND NOT xSenseExtend, PT := tSensorTimeout);

IF xSenseRetract AND xSenseExtend THEN
	(* 两端同时有信号：传感器短路、磁环位置错或机械卡在中间，姿态不可信 *)
	xPositionKnown := FALSE;
	stStatus.lrPosition := lrLastKnown;
	stStatus.xError := TRUE; stStatus.udiErrorID := 3003;
ELSIF xSenseExtend THEN
	xPositionKnown := TRUE; lrLastKnown := 1.0; stStatus.lrPosition := 1.0;
ELSIF xSenseRetract THEN
	xPositionKnown := TRUE; lrLastKnown := 0.0; stStatus.lrPosition := 0.0;
ELSE
	(* 两端都没有信号：保持最后姿态；从未确立过则 xReady 一直为 FALSE *)
	stStatus.lrPosition := lrLastKnown;
	IF tonNoSensor.Q AND NOT stStatus.xError THEN
		xPositionKnown := FALSE;
		stStatus.xError := TRUE; stStatus.udiErrorID := 3004;
	END_IF
END_IF

(* ===== 3. 命令接收与保位判定 ===== *)
IF NOT xUseReal THEN
	(* 未接管：不驱动阀，也不发布就绪，避免被上层当成可用设备 *)
	xCmdValid := FALSE; xTravelling := FALSE; udiLastID := 0;
	stStatus.xReady := FALSE; stStatus.xBusy := FALSE; stStatus.xActive := FALSE;
	stStatus.udiAcceptedID := 0; stStatus.udiCompletedID := 0;
ELSIF NOT xEnable OR stStatus.xError OR xFaultHold THEN
	(* 故障或整机故障保持时阀失电，不带错误继续动作 *)
	xCmdValid := FALSE; xTravelling := FALSE;
	stStatus.xReady := FALSE; stStatus.xBusy := FALSE; stStatus.xActive := FALSE;
ELSE
	stStatus.xReady := xEnable AND xPositionKnown;

	(* 新序号即新命令；姿态未确立时不接受，防止朝未知状态动作 *)
	IF (stCommand.udiID <> 0) AND (stCommand.udiID <> udiLastID)
		AND xEnable AND xPositionKnown AND NOT stStatus.xBusy THEN
		udiLastID := stCommand.udiID;
		stStatus.udiAcceptedID := udiLastID; stStatus.udiCompletedID := 0;
		CASE stCommand.eAction OF
		E_DeviceAction.Position:
			IF (stCommand.lrTarget < stConfig.lrMinPosition - 0.01)
				OR (stCommand.lrTarget > stConfig.lrMaxPosition + 0.01) THEN
				stStatus.xError := TRUE; stStatus.udiErrorID := 2001;
				xCmdValid := FALSE;
			ELSE
				xCmdExtend := stCommand.lrTarget > 0.5;
				xCmdValid := TRUE;
				xTravelling := TRUE;
				stStatus.xBusy := TRUE;
			END_IF
		E_DeviceAction.Stop, E_DeviceAction.None:
			xCmdValid := FALSE; xTravelling := FALSE;
			stStatus.udiAcceptedID := 0; stStatus.udiCompletedID := 0;
			udiLastID := 0;
		ELSE
			(* 气缸没有连续运行、点动和回零，明确报错而不是静默不动 *)
			stStatus.xError := TRUE; stStatus.udiErrorID := 2001;
			xCmdValid := FALSE;
		END_CASE
	END_IF

	(* 命令被撤销或失能：立即取消保位，阀随之失电 *)
	IF (stCommand.eAction = E_DeviceAction.Stop) OR (stCommand.eAction = E_DeviceAction.None)
		OR NOT xEnable THEN
		xCmdValid := FALSE; xTravelling := FALSE;
		stStatus.xBusy := FALSE;
	END_IF

	(* 到位判定：姿态已知且与命令期望的端点一致即算完成 *)
	IF xCmdValid AND xPositionKnown THEN
		IF (xCmdExtend AND (stStatus.lrPosition > 0.5))
			OR ((NOT xCmdExtend) AND (stStatus.lrPosition < 0.5)) THEN
			IF xTravelling THEN stStatus.udiCompletedID := udiLastID; END_IF
			xTravelling := FALSE;
			stStatus.xBusy := FALSE;
		END_IF
	END_IF
END_IF

(* ===== 4. 到位超时 ===== *)
tonTravel(IN := xUseReal AND xTravelling AND xCmdValid, PT := tTravelTimeout);
IF tonTravel.Q AND NOT stStatus.xError THEN
	stStatus.xError := TRUE; stStatus.udiErrorID := 3005;
	stStatus.xBusy := FALSE;
	xTravelling := FALSE;
END_IF

(* ===== 5. 阀输出：按保位命令持续输出，不是只在动作过程中输出 ===== *)
xValve := FALSE;
xValve2 := FALSE;
IF xCmdValid AND xUseReal AND NOT stStatus.xError AND NOT xFaultHold THEN
	xValve := xCmdExtend;
	IF xUseSecond THEN xValve2 := xCmdExtend; END_IF
END_IF
IF xInvertValve THEN xValve := NOT xValve; END_IF
IF xInvertValve AND xUseSecond THEN xValve2 := NOT xValve2; END_IF

(* ===== 6. 收尾 ===== *)
stStatus.xReady := stStatus.xReady AND xUseReal AND NOT stStatus.xError;
stStatus.xActive := xCmdValid;
(* 气缸没有回零动作，用“姿态已确立”代替，供整机统计已接管设备是否可信 *)
stStatus.xHomed := xUseReal AND xPositionKnown;

END_FUNCTION_BLOCK

